(* IEC 61131-3 sources: plc-st-coding-agent/progress/evidence/f14_v3_parallel_20261112/jobs/codex_minimax-m27 (part 2) *)

(* ---- public-hard-05.raw_candidate_01.st ---- *)
FUNCTION_BLOCK MechanicalArmControl
VAR_INPUT
    ManualMode      : BOOL;
    SingleStepMode  : BOOL;
    SingleCycleMode : BOOL;
    ContinuousMode  : BOOL;
    EmergencyStop   : BOOL;
    Start           : BOOL;
    DownButton      : BOOL;
    UpButton        : BOOL;
    LeftButton      : BOOL;
    RightButton     : BOOL;
    GripButton      : BOOL;
    ReleaseButton   : BOOL;
    DownLimitSwitch     : BOOL;
    UpLimitSwitch       : BOOL;
    LeftLimitSwitch     : BOOL;
    RightLimitSwitch    : BOOL;
    GripLimitSwitch     : BOOL;
    ReleaseLimitSwitch  : BOOL;
END_VAR

VAR_OUTPUT
    MoveDown        : BOOL;
    MoveUp          : BOOL;
    MoveLeft        : BOOL;
    MoveRight       : BOOL;
    ActivateGrip    : BOOL;
    ActivateRelease : BOOL;
END_VAR

VAR
    stepNumber       : INT := 0;
    startRisingEdge  : BOOL;
    lastStart        : BOOL := FALSE;
    actionInProgress : BOOL := FALSE;
END_VAR

// Edge detection for Start button
startRisingEdge := Start AND NOT lastStart;
lastStart := Start;

// Emergency stop: highest priority, resets all outputs and state
IF NOT EmergencyStop THEN
    MoveDown        := FALSE;
    MoveUp          := FALSE;
    MoveLeft        := FALSE;
    MoveRight       := FALSE;
    ActivateGrip    := FALSE;
    ActivateRelease := FALSE;
    stepNumber      := 0;
    actionInProgress := FALSE;
ELSE
    // Manual mode control
    IF ManualMode THEN
        MoveDown        := DownButton AND NOT DownLimitSwitch;
        MoveUp          := UpButton AND NOT UpLimitSwitch;
        MoveLeft        := LeftButton AND NOT LeftLimitSwitch;
        MoveRight       := RightButton AND NOT RightLimitSwitch;
        ActivateGrip    := GripButton AND NOT GripLimitSwitch;
        ActivateRelease := ReleaseButton AND NOT ReleaseLimitSwitch;
        stepNumber      := 0;
        actionInProgress := FALSE;

    // Single step mode: Start button advances through steps
    ELSIF SingleStepMode THEN
        IF startRisingEdge AND NOT actionInProgress THEN
            stepNumber := stepNumber + 1;
        END_IF;

        CASE stepNumber OF
            1:
                MoveDown := TRUE;
                actionInProgress := TRUE;
                IF DownLimitSwitch THEN
                    MoveDown := FALSE;
                    actionInProgress := FALSE;
                END_IF;
            2:
                ActivateGrip := TRUE;
                actionInProgress := TRUE;
                IF GripLimitSwitch THEN
                    ActivateGrip := FALSE;
                    actionInProgress := FALSE;
                END_IF;
            3:
                MoveUp := TRUE;
                actionInProgress := TRUE;
                IF UpLimitSwitch THEN
                    MoveUp := FALSE;
                    actionInProgress := FALSE;
                END_IF;
            4:
                MoveRight := TRUE;
                actionInProgress := TRUE;
                IF RightLimitSwitch THEN
                    MoveRight := FALSE;
                    actionInProgress := FALSE;
                END_IF;
            5:
                MoveDown := TRUE;
                actionInProgress := TRUE;
                IF DownLimitSwitch THEN
                    MoveDown := FALSE;
                    actionInProgress := FALSE;
                END_IF;
            6:
                ActivateRelease := TRUE;
                actionInProgress := TRUE;
                IF ReleaseLimitSwitch THEN
                    ActivateRelease := FALSE;
                    actionInProgress := FALSE;
                END_IF;
            7:
                MoveUp := TRUE;
                actionInProgress := TRUE;
                IF UpLimitSwitch THEN
                    MoveUp := FALSE;
                    actionInProgress := FALSE;
                END_IF;
            8:
                MoveLeft := TRUE;
                actionInProgress := TRUE;
                IF LeftLimitSwitch THEN
                    MoveLeft := FALSE;
                    actionInProgress := FALSE;
                END_IF;
        END_CASE;

        IF stepNumber > 8 THEN
            stepNumber := 0;
        END_IF;

    // Single cycle mode: executes full cycle once then stops
    ELSIF SingleCycleMode THEN
        IF startRisingEdge THEN
            stepNumber := 1;
            actionInProgress := FALSE;
        END_IF;

        CASE stepNumber OF
            1:
                MoveDown := TRUE;
                actionInProgress := TRUE;
                IF DownLimitSwitch THEN
                    MoveDown := FALSE;
                    actionInProgress := FALSE;
                    stepNumber := 2;
                END_IF;
            2:
                ActivateGrip := TRUE;
                actionInProgress := TRUE;
                IF GripLimitSwitch THEN
                    ActivateGrip := FALSE;
                    actionInProgress := FALSE;
                    stepNumber := 3;
                END_IF;
            3:
                MoveUp := TRUE;
                actionInProgress := TRUE;
                IF UpLimitSwitch THEN
                    MoveUp := FALSE;
                    actionInProgress := FALSE;
                    stepNumber := 4;
                END_IF;
            4:
                MoveRight := TRUE;
                actionInProgress := TRUE;
                IF RightLimitSwitch THEN
                    MoveRight := FALSE;
                    actionInProgress := FALSE;
                    stepNumber := 5;
                END_IF;
            5:
                MoveDown := TRUE;
                actionInProgress := TRUE;
                IF DownLimitSwitch THEN
                    MoveDown := FALSE;
                    actionInProgress := FALSE;
                    stepNumber := 6;
                END_IF;
            6:
                ActivateRelease := TRUE;
                actionInProgress := TRUE;
                IF ReleaseLimitSwitch THEN
                    ActivateRelease := FALSE;
                    actionInProgress := FALSE;
                    stepNumber := 7;
                END_IF;
            7:
                MoveUp := TRUE;
                actionInProgress := TRUE;
                IF UpLimitSwitch THEN
                    MoveUp := FALSE;
                    actionInProgress := FALSE;
                    stepNumber := 8;
                END_IF;
            8:
                MoveLeft := TRUE;
                actionInProgress := TRUE;
                IF LeftLimitSwitch THEN
                    MoveLeft := FALSE;
                    actionInProgress := FALSE;
                    stepNumber := 0;
                END_IF;
        END_CASE;

    // Continuous mode: executes full cycle repeatedly
    ELSIF ContinuousMode THEN
        IF startRisingEdge THEN
            stepNumber := 1;
            actionInProgress := FALSE;
        END_IF;

        CASE stepNumber OF
            1:
                MoveDown := TRUE;
                actionInProgress := TRUE;
                IF DownLimitSwitch THEN
                    MoveDown := FALSE;
                    actionInProgress := FALSE;
                    stepNumber := 2;
                END_IF;
            2:
                ActivateGrip := TRUE;
                actionInProgress := TRUE;
                IF GripLimitSwitch THEN
                    ActivateGrip := FALSE;
                    actionInProgress := FALSE;
                    stepNumber := 3;
                END_IF;
            3:
                MoveUp := TRUE;
                actionInProgress := TRUE;
                IF UpLimitSwitch THEN
                    MoveUp := FALSE;
                    actionInProgress := FALSE;
                    stepNumber := 4;
                END_IF;
            4:
                MoveRight := TRUE;
                actionInProgress := TRUE;
                IF RightLimitSwitch THEN
                    MoveRight := FALSE;
                    actionInProgress := FALSE;
                    stepNumber := 5;
                END_IF;
            5:
                MoveDown := TRUE;
                actionInProgress := TRUE;
                IF DownLimitSwitch THEN
                    MoveDown := FALSE;
                    actionInProgress := FALSE;
                    stepNumber := 6;
                END_IF;
            6:
                ActivateRelease := TRUE;
                actionInProgress := TRUE;
                IF ReleaseLimitSwitch THEN
                    ActivateRelease := FALSE;
                    actionInProgress := FALSE;
                    stepNumber := 7;
                END_IF;
            7:
                MoveUp := TRUE;
                actionInProgress := TRUE;
                IF UpLimitSwitch THEN
                    MoveUp := FALSE;
                    actionInProgress := FALSE;
                    stepNumber := 8;
                END_IF;
            8:
                MoveLeft := TRUE;
                actionInProgress := TRUE;
                IF LeftLimitSwitch THEN
                    MoveLeft := FALSE;
                    actionInProgress := FALSE;
                    stepNumber := 1;
                END_IF;
        END_CASE;
    END_IF;
END_IF;
END_FUNCTION_BLOCK

(* ---- public-hard-05.raw_candidate_02.st ---- *)
FUNCTION_BLOCK MechanicalArmControl
VAR_INPUT
    ManualMode      : BOOL;
    SingleStepMode  : BOOL;
    SingleCycleMode : BOOL;
    ContinuousMode  : BOOL;
    EmergencyStop   : BOOL;
    Start           : BOOL;
    DownButton      : BOOL;
    UpButton        : BOOL;
    LeftButton      : BOOL;
    RightButton     : BOOL;
    GripButton      : BOOL;
    ReleaseButton   : BOOL;
    DownLimitSwitch     : BOOL;
    UpLimitSwitch       : BOOL;
    LeftLimitSwitch     : BOOL;
    RightLimitSwitch    : BOOL;
    GripLimitSwitch     : BOOL;
    ReleaseLimitSwitch  : BOOL;
END_VAR

VAR_OUTPUT
    MoveDown        : BOOL;
    MoveUp          : BOOL;
    MoveLeft        : BOOL;
    MoveRight       : BOOL;
    ActivateGrip    : BOOL;
    ActivateRelease : BOOL;
END_VAR

VAR
    stepNumber       : INT := 0;
    startRisingEdge  : BOOL;
    lastStart        : BOOL := FALSE;
    actionInProgress : BOOL := FALSE;
END_VAR

startRisingEdge := Start AND NOT lastStart;
lastStart := Start;

IF NOT EmergencyStop THEN
    MoveDown        := FALSE;
    MoveUp          := FALSE;
    MoveLeft        := FALSE;
    MoveRight       := FALSE;
    ActivateGrip    := FALSE;
    ActivateRelease := FALSE;
    stepNumber      := 0;
    actionInProgress := FALSE;
ELSE
    IF ManualMode THEN
        IF DownButton AND UpButton THEN
            MoveDown := FALSE;
            MoveUp := FALSE;
        ELSE
            MoveDown := DownButton AND NOT DownLimitSwitch;
            MoveUp := UpButton AND NOT UpLimitSwitch;
        END_IF;
        IF LeftButton AND RightButton THEN
            MoveLeft := FALSE;
            MoveRight := FALSE;
        ELSE
            MoveLeft := LeftButton AND NOT LeftLimitSwitch;
            MoveRight := RightButton AND NOT RightLimitSwitch;
        END_IF;
        ActivateGrip := GripButton AND NOT GripLimitSwitch;
        ActivateRelease := ReleaseButton AND NOT ReleaseLimitSwitch;
        stepNumber := 0;
        actionInProgress := FALSE;

    ELSIF SingleStepMode THEN
        IF startRisingEdge AND NOT actionInProgress THEN
            stepNumber := stepNumber + 1;
        END_IF;

        IF stepNumber = 0 THEN
            actionInProgress := FALSE;
        END_IF;

        CASE stepNumber OF
            1:
                MoveDown := TRUE;
                actionInProgress := TRUE;
                IF DownLimitSwitch THEN
                    MoveDown := FALSE;
                    actionInProgress := FALSE;
                END_IF;
            2:
                ActivateGrip := TRUE;
                actionInProgress := TRUE;
                IF GripLimitSwitch THEN
                    ActivateGrip := FALSE;
                    actionInProgress := FALSE;
                END_IF;
            3:
                MoveUp := TRUE;
                actionInProgress := TRUE;
                IF UpLimitSwitch THEN
                    MoveUp := FALSE;
                    actionInProgress := FALSE;
                END_IF;
            4:
                MoveRight := TRUE;
                actionInProgress := TRUE;
                IF RightLimitSwitch THEN
                    MoveRight := FALSE;
                    actionInProgress := FALSE;
                END_IF;
            5:
                MoveDown := TRUE;
                actionInProgress := TRUE;
                IF DownLimitSwitch THEN
                    MoveDown := FALSE;
                    actionInProgress := FALSE;
                END_IF;
            6:
                ActivateRelease := TRUE;
                actionInProgress := TRUE;
                IF ReleaseLimitSwitch THEN
                    ActivateRelease := FALSE;
                    actionInProgress := FALSE;
                END_IF;
            7:
                MoveUp := TRUE;
                actionInProgress := TRUE;
                IF UpLimitSwitch THEN
                    MoveUp := FALSE;
                    actionInProgress := FALSE;
                END_IF;
            8:
                MoveLeft := TRUE;
                actionInProgress := TRUE;
                IF LeftLimitSwitch THEN
                    MoveLeft := FALSE;
                    actionInProgress := FALSE;
                END_IF;
        END_CASE;

        IF stepNumber > 8 THEN
            stepNumber := 0;
        END_IF;

    ELSIF SingleCycleMode THEN
        IF startRisingEdge THEN
            stepNumber := 1;
            actionInProgress := FALSE;
        END_IF;

        IF stepNumber = 0 THEN
            actionInProgress := FALSE;
        END_IF;

        CASE stepNumber OF
            1:
                MoveDown := TRUE;
                actionInProgress := TRUE;
                IF DownLimitSwitch THEN
                    MoveDown := FALSE;
                    actionInProgress := FALSE;
                    stepNumber := 2;
                END_IF;
            2:
                ActivateGrip := TRUE;
                actionInProgress := TRUE;
                IF GripLimitSwitch THEN
                    ActivateGrip := FALSE;
                    actionInProgress := FALSE;
                    stepNumber := 3;
                END_IF;
            3:
                MoveUp := TRUE;
                actionInProgress := TRUE;
                IF UpLimitSwitch THEN
                    MoveUp := FALSE;
                    actionInProgress := FALSE;
                    stepNumber := 4;
                END_IF;
            4:
                MoveRight := TRUE;
                actionInProgress := TRUE;
                IF RightLimitSwitch THEN
                    MoveRight := FALSE;
                    actionInProgress := FALSE;
                    stepNumber := 5;
                END_IF;
            5:
                MoveDown := TRUE;
                actionInProgress := TRUE;
                IF DownLimitSwitch THEN
                    MoveDown := FALSE;
                    actionInProgress := FALSE;
                    stepNumber := 6;
                END_IF;
            6:
                ActivateRelease := TRUE;
                actionInProgress := TRUE;
                IF ReleaseLimitSwitch THEN
                    ActivateRelease := FALSE;
                    actionInProgress := FALSE;
                    stepNumber := 7;
                END_IF;
            7:
                MoveUp := TRUE;
                actionInProgress := TRUE;
                IF UpLimitSwitch THEN
                    MoveUp := FALSE;
                    actionInProgress := FALSE;
                    stepNumber := 8;
                END_IF;
            8:
                MoveLeft := TRUE;
                actionInProgress := TRUE;
                IF LeftLimitSwitch THEN
                    MoveLeft := FALSE;
                    actionInProgress := FALSE;
                    stepNumber := 0;
                END_IF;
        END_CASE;

    ELSIF ContinuousMode THEN
        IF startRisingEdge THEN
            stepNumber := 1;
            actionInProgress := FALSE;
        END_IF;

        IF stepNumber = 0 THEN
            actionInProgress := FALSE;
        END_IF;

        CASE stepNumber OF
            1:
                MoveDown := TRUE;
                actionInProgress := TRUE;
                IF DownLimitSwitch THEN
                    MoveDown := FALSE;
                    actionInProgress := FALSE;
                    stepNumber := 2;
                END_IF;
            2:
                ActivateGrip := TRUE;
                actionInProgress := TRUE;
                IF GripLimitSwitch THEN
                    ActivateGrip := FALSE;
                    actionInProgress := FALSE;
                    stepNumber := 3;
                END_IF;
            3:
                MoveUp := TRUE;
                actionInProgress := TRUE;
                IF UpLimitSwitch THEN
                    MoveUp := FALSE;
                    actionInProgress := FALSE;
                    stepNumber := 4;
                END_IF;
            4:
                MoveRight := TRUE;
                actionInProgress := TRUE;
                IF RightLimitSwitch THEN
                    MoveRight := FALSE;
                    actionInProgress := FALSE;
                    stepNumber := 5;
                END_IF;
            5:
                MoveDown := TRUE;
                actionInProgress := TRUE;
                IF DownLimitSwitch THEN
                    MoveDown := FALSE;
                    actionInProgress := FALSE;
                    stepNumber := 6;
                END_IF;
            6:
                ActivateRelease := TRUE;
                actionInProgress := TRUE;
                IF ReleaseLimitSwitch THEN
                    ActivateRelease := FALSE;
                    actionInProgress := FALSE;
                    stepNumber := 7;
                END_IF;
            7:
                MoveUp := TRUE;
                actionInProgress := TRUE;
                IF UpLimitSwitch THEN
                    MoveUp := FALSE;
                    actionInProgress := FALSE;
                    stepNumber := 8;
                END_IF;
            8:
                MoveLeft := TRUE;
                actionInProgress := TRUE;
                IF LeftLimitSwitch THEN
                    MoveLeft := FALSE;
                    actionInProgress := FALSE;
                    stepNumber := 1;
                END_IF;
        END_CASE;
    END_IF;
END_IF;
END_FUNCTION_BLOCK

(* ---- public-hard-06.candidate_01.st ---- *)
TYPE ProductState : (
    Idle := 0,
    AtFeed := 1,
    AtWash := 2,
    AtWeight := 3,
    AtFiring := 4,
    AtOutput := 5,
    Rejected := 6
);
END_TYPE;

FUNCTION_BLOCK ProductionControl
VAR_INPUT
    Mode : BOOL;
    ForwardButton : BOOL;
    ReverseButton : BOOL;
    SensorFeed : BOOL;
    SensorWash : BOOL;
    SensorWeight : BOOL;
    SensorFiring : BOOL;
    SensorOutput : BOOL;
    washComplete : BOOL;
    weightComplete : BOOL;
    weight : REAL;
    firingComplete : BOOL;
END_VAR

VAR_OUTPUT
    MotorForward : BOOL := FALSE;
    MotorReverse : BOOL := FALSE;
    kick : BOOL := FALSE;
    CompletionLight : BOOL := FALSE;
    firingTemp : REAL := 0.0;
END_VAR

VAR
    currentState : ProductState := Idle;
    prevSensorFeed : BOOL := FALSE;
    prevSensorWash : BOOL := FALSE;
    prevSensorWeight : BOOL := FALSE;
    prevSensorFiring : BOOL := FALSE;
    prevSensorOutput : BOOL := FALSE;
END_VAR

IF currentState = Idle THEN
    MotorForward := FALSE;
    MotorReverse := FALSE;
    kick := FALSE;
    CompletionLight := FALSE;
    firingTemp := 0.0;
END_IF;

IF Mode = FALSE THEN
    MotorForward := ForwardButton;
    MotorReverse := ReverseButton AND NOT ForwardButton;
    MotorReverse := MotorReverse;
ELSE
    MotorReverse := FALSE;

    IF currentState = Idle THEN
        IF SensorFeed AND NOT prevSensorFeed THEN
            currentState := AtFeed;
            MotorForward := TRUE;
        END_IF;

    ELSIF currentState = AtFeed THEN
        MotorForward := TRUE;
        IF SensorWash AND NOT prevSensorWash THEN
            currentState := AtWash;
            MotorForward := FALSE;
        END_IF;

    ELSIF currentState = AtWash THEN
        MotorForward := FALSE;
        IF washComplete THEN
            currentState := AtWeight;
            MotorForward := TRUE;
        END_IF;

    ELSIF currentState = AtWeight THEN
        MotorForward := FALSE;
        IF weightComplete THEN
            IF weight < 100.0 OR weight > 200.0 THEN
                kick := TRUE;
                currentState := Rejected;
                MotorForward := TRUE;
            ELSE
                firingTemp := 500.0 + (weight - 100.0) * 0.5;
                currentState := AtFiring;
                MotorForward := TRUE;
            END_IF;
        END_IF;

    ELSIF currentState = AtFiring THEN
        MotorForward := FALSE;
        IF firingComplete THEN
            currentState := AtOutput;
            MotorForward := FALSE;
            CompletionLight := TRUE;
        END_IF;

    ELSIF currentState = AtOutput THEN
        MotorForward := FALSE;
        CompletionLight := SensorOutput;
        IF NOT SensorOutput AND prevSensorOutput THEN
            currentState := Idle;
            CompletionLight := FALSE;
        END_IF;

    ELSIF currentState = Rejected THEN
        MotorForward := TRUE;
        kick := SensorWeight;
        IF NOT SensorWeight AND prevSensorWeight THEN
            currentState := Idle;
            kick := FALSE;
        END_IF;

    END_IF;
END_IF;

prevSensorFeed := SensorFeed;
prevSensorWash := SensorWash;
prevSensorWeight := SensorWeight;
prevSensorFiring := SensorFiring;
prevSensorOutput := SensorOutput;

END_FUNCTION_BLOCK

(* ---- public-hard-06.candidate_02.st ---- *)
TYPE ProductState : (
    Idle := 0,
    AtFeed := 1,
    AtWash := 2,
    AtWeight := 3,
    AtFiring := 4,
    AtOutput := 5,
    Rejected := 6
);
END_TYPE;

TYPE ModeType : (Manual := 0, Auto := 1, Sequence := 2);
END_TYPE;

FUNCTION_BLOCK ProductionControl
VAR_INPUT
    Mode : BOOL;
    ForwardButton : BOOL;
    ReverseButton : BOOL;
    SensorFeed : BOOL;
    SensorWash : BOOL;
    SensorWeight : BOOL;
    SensorFiring : BOOL;
    SensorOutput : BOOL;
    washComplete : BOOL;
    weightComplete : BOOL;
    weight : REAL;
    firingComplete : BOOL;
END_VAR

VAR_OUTPUT
    MotorForward : BOOL := FALSE;
    MotorReverse : BOOL := FALSE;
    kick : BOOL := FALSE;
    CompletionLight : BOOL := FALSE;
    firingTemp : REAL := 0.0;
END_VAR

VAR
    currentState : ProductState := Idle;
    prevSensorFeed : BOOL := FALSE;
    prevSensorWash : BOOL := FALSE;
    prevSensorWeight : BOOL := FALSE;
    prevSensorFiring : BOOL := FALSE;
    prevSensorOutput : BOOL := FALSE;
    prevWashComplete : BOOL := FALSE;
    prevWeightComplete : BOOL := FALSE;
    prevFiringComplete : BOOL := FALSE;
END_VAR

IF currentState = Idle THEN
    MotorForward := FALSE;
    MotorReverse := FALSE;
    kick := FALSE;
    CompletionLight := FALSE;
    firingTemp := 0.0;
END_IF;

IF Mode = FALSE THEN
    MotorForward := ForwardButton;
    MotorReverse := ReverseButton AND NOT ForwardButton;
ELSE
    MotorReverse := FALSE;

    IF currentState = Idle THEN
        IF SensorFeed AND NOT prevSensorFeed THEN
            currentState := AtFeed;
            MotorForward := TRUE;
        END_IF;

    ELSIF currentState = AtFeed THEN
        MotorForward := TRUE;
        IF SensorWash AND NOT prevSensorWash THEN
            currentState := AtWash;
            MotorForward := FALSE;
        END_IF;

    ELSIF currentState = AtWash THEN
        MotorForward := FALSE;
        IF washComplete AND NOT prevWashComplete THEN
            currentState := AtWeight;
            MotorForward := TRUE;
        END_IF;

    ELSIF currentState = AtWeight THEN
        MotorForward := FALSE;
        IF weightComplete AND NOT prevWeightComplete THEN
            IF weight < 100.0 OR weight > 200.0 THEN
                kick := TRUE;
                currentState := Rejected;
            ELSE
                firingTemp := 500.0 + (weight - 100.0) * 0.5;
                currentState := AtFiring;
            END_IF;
        END_IF;

    ELSIF currentState = AtFiring THEN
        MotorForward := FALSE;
        IF firingComplete AND NOT prevFiringComplete THEN
            currentState := AtOutput;
            CompletionLight := TRUE;
        END_IF;

    ELSIF currentState = AtOutput THEN
        MotorForward := FALSE;
        CompletionLight := SensorOutput;
        IF NOT SensorOutput AND prevSensorOutput THEN
            currentState := Idle;
            CompletionLight := FALSE;
        END_IF;

    ELSIF currentState = Rejected THEN
        MotorForward := FALSE;
        kick := SensorWeight;
        IF NOT SensorWeight AND prevSensorWeight THEN
            currentState := Idle;
            kick := FALSE;
        END_IF;

    END_IF;
END_IF;

prevSensorFeed := SensorFeed;
prevSensorWash := SensorWash;
prevSensorWeight := SensorWeight;
prevSensorFiring := SensorFiring;
prevSensorOutput := SensorOutput;
prevWashComplete := washComplete;
prevWeightComplete := weightComplete;
prevFiringComplete := firingComplete;

END_FUNCTION_BLOCK

(* ---- public-hard-06.raw_candidate_01.st ---- *)
TYPE ProductState : (
    Idle := 0,
    AtFeed := 1,
    AtWash := 2,
    AtWeight := 3,
    AtFiring := 4,
    AtOutput := 5,
    Rejected := 6
);
END_TYPE

FUNCTION_BLOCK ProductionControl
VAR_INPUT
    Mode : BOOL;
    ForwardButton : BOOL;
    ReverseButton : BOOL;
    SensorFeed : BOOL;
    SensorWash : BOOL;
    SensorWeight : BOOL;
    SensorFiring : BOOL;
    SensorOutput : BOOL;
    washComplete : BOOL;
    weightComplete : BOOL;
    weight : REAL;
    firingComplete : BOOL;
END_VAR

VAR_OUTPUT
    MotorForward : BOOL := FALSE;
    MotorReverse : BOOL := FALSE;
    kick : BOOL := FALSE;
    CompletionLight : BOOL := FALSE;
    firingTemp : REAL := 0.0;
END_VAR

VAR
    currentState : ProductState := Idle;
    prevSensorFeed : BOOL := FALSE;
    prevSensorWash : BOOL := FALSE;
    prevSensorWeight : BOOL := FALSE;
    prevSensorFiring : BOOL := FALSE;
    prevSensorOutput : BOOL := FALSE;
END_VAR

IF currentState = Idle THEN
    MotorForward := FALSE;
    MotorReverse := FALSE;
    kick := FALSE;
    CompletionLight := FALSE;
    firingTemp := 0.0;
END_IF

IF Mode = FALSE THEN
    MotorForward := ForwardButton;
    MotorReverse := ReverseButton AND NOT ForwardButton;
    MotorReverse := MotorReverse;
ELSE
    MotorReverse := FALSE;

    IF currentState = Idle THEN
        IF SensorFeed AND NOT prevSensorFeed THEN
            currentState := AtFeed;
            MotorForward := TRUE;
        END_IF

    ELSIF currentState = AtFeed THEN
        MotorForward := TRUE;
        IF SensorWash AND NOT prevSensorWash THEN
            currentState := AtWash;
            MotorForward := FALSE;
        END_IF

    ELSIF currentState = AtWash THEN
        MotorForward := FALSE;
        IF washComplete THEN
            currentState := AtWeight;
            MotorForward := TRUE;
        END_IF

    ELSIF currentState = AtWeight THEN
        MotorForward := FALSE;
        IF weightComplete THEN
            IF weight < 100.0 OR weight > 200.0 THEN
                kick := TRUE;
                currentState := Rejected;
                MotorForward := TRUE;
            ELSE
                firingTemp := 500.0 + (weight - 100.0) * 0.5;
                currentState := AtFiring;
                MotorForward := TRUE;
            END_IF;
        END_IF

    ELSIF currentState = AtFiring THEN
        MotorForward := FALSE;
        IF firingComplete THEN
            currentState := AtOutput;
            MotorForward := FALSE;
            CompletionLight := TRUE;
        END_IF

    ELSIF currentState = AtOutput THEN
        MotorForward := FALSE;
        CompletionLight := SensorOutput;
        IF NOT SensorOutput AND prevSensorOutput THEN
            currentState := Idle;
            CompletionLight := FALSE;
        END_IF

    ELSIF currentState = Rejected THEN
        MotorForward := TRUE;
        kick := SensorWeight;
        IF NOT SensorWeight AND prevSensorWeight THEN
            currentState := Idle;
            kick := FALSE;
        END_IF

    END_IF
END_IF

prevSensorFeed := SensorFeed;
prevSensorWash := SensorWash;
prevSensorWeight := SensorWeight;
prevSensorFiring := SensorFiring;
prevSensorOutput := SensorOutput;

END_FUNCTION_BLOCK

(* ---- public-hard-06.raw_candidate_02.st ---- *)
TYPE ProductState : (
    Idle := 0,
    AtFeed := 1,
    AtWash := 2,
    AtWeight := 3,
    AtFiring := 4,
    AtOutput := 5,
    Rejected := 6
);
END_TYPE

TYPE ModeType : (Manual := 0, Auto := 1, Sequence := 2);
END_TYPE

FUNCTION_BLOCK ProductionControl
VAR_INPUT
    Mode : BOOL;
    ForwardButton : BOOL;
    ReverseButton : BOOL;
    SensorFeed : BOOL;
    SensorWash : BOOL;
    SensorWeight : BOOL;
    SensorFiring : BOOL;
    SensorOutput : BOOL;
    washComplete : BOOL;
    weightComplete : BOOL;
    weight : REAL;
    firingComplete : BOOL;
END_VAR

VAR_OUTPUT
    MotorForward : BOOL := FALSE;
    MotorReverse : BOOL := FALSE;
    kick : BOOL := FALSE;
    CompletionLight : BOOL := FALSE;
    firingTemp : REAL := 0.0;
END_VAR

VAR
    currentState : ProductState := Idle;
    prevSensorFeed : BOOL := FALSE;
    prevSensorWash : BOOL := FALSE;
    prevSensorWeight : BOOL := FALSE;
    prevSensorFiring : BOOL := FALSE;
    prevSensorOutput : BOOL := FALSE;
    prevWashComplete : BOOL := FALSE;
    prevWeightComplete : BOOL := FALSE;
    prevFiringComplete : BOOL := FALSE;
END_VAR

IF currentState = Idle THEN
    MotorForward := FALSE;
    MotorReverse := FALSE;
    kick := FALSE;
    CompletionLight := FALSE;
    firingTemp := 0.0;
END_IF;

IF Mode = FALSE THEN
    MotorForward := ForwardButton;
    MotorReverse := ReverseButton AND NOT ForwardButton;
ELSE
    MotorReverse := FALSE;

    IF currentState = Idle THEN
        IF SensorFeed AND NOT prevSensorFeed THEN
            currentState := AtFeed;
            MotorForward := TRUE;
        END_IF;

    ELSIF currentState = AtFeed THEN
        MotorForward := TRUE;
        IF SensorWash AND NOT prevSensorWash THEN
            currentState := AtWash;
            MotorForward := FALSE;
        END_IF;

    ELSIF currentState = AtWash THEN
        MotorForward := FALSE;
        IF washComplete AND NOT prevWashComplete THEN
            currentState := AtWeight;
            MotorForward := TRUE;
        END_IF;

    ELSIF currentState = AtWeight THEN
        MotorForward := FALSE;
        IF weightComplete AND NOT prevWeightComplete THEN
            IF weight < 100.0 OR weight > 200.0 THEN
                kick := TRUE;
                currentState := Rejected;
            ELSE
                firingTemp := 500.0 + (weight - 100.0) * 0.5;
                currentState := AtFiring;
            END_IF;
        END_IF;

    ELSIF currentState = AtFiring THEN
        MotorForward := FALSE;
        IF firingComplete AND NOT prevFiringComplete THEN
            currentState := AtOutput;
            CompletionLight := TRUE;
        END_IF;

    ELSIF currentState = AtOutput THEN
        MotorForward := FALSE;
        CompletionLight := SensorOutput;
        IF NOT SensorOutput AND prevSensorOutput THEN
            currentState := Idle;
            CompletionLight := FALSE;
        END_IF;

    ELSIF currentState = Rejected THEN
        MotorForward := FALSE;
        kick := SensorWeight;
        IF NOT SensorWeight AND prevSensorWeight THEN
            currentState := Idle;
            kick := FALSE;
        END_IF;

    END_IF;
END_IF;

prevSensorFeed := SensorFeed;
prevSensorWash := SensorWash;
prevSensorWeight := SensorWeight;
prevSensorFiring := SensorFiring;
prevSensorOutput := SensorOutput;
prevWashComplete := washComplete;
prevWeightComplete := weightComplete;
prevFiringComplete := firingComplete;

END_FUNCTION_BLOCK

(* ---- public-medium-01.candidate_01.st ---- *)
FUNCTION_BLOCK FB_PumpControl
VAR
    i : INT;
    sortedIndices : ARRAY[1..5] OF INT;
    temp : INT;
    j : INT;
END_VAR

    // Stop button has highest priority
    IF stop THEN
        FOR i := 1 TO 5 DO
            pumpGroup[i].RunComd := FALSE;
        END_FOR;
        RETURN;
    END_IF;

    // Start button applies mode-specific logic
    IF start THEN
        IF NOT mode THEN
            // Manual mode - run pumps where selection is TRUE
            FOR i := 1 TO 5 DO
                pumpGroup[i].RunComd := pumpGroup[i].selection;
            END_FOR;
        ELSE
            // Automatic mode - select 3 pumps with highest priority
            FOR i := 1 TO 5 DO
                sortedIndices[i] := i;
            END_FOR;

            // Bubble sort by priority (descending)
            FOR i := 1 TO 4 DO
                FOR j := i + 1 TO 5 DO
                    IF pumpGroup[sortedIndices[j]].priority > pumpGroup[sortedIndices[i]].priority THEN
                        temp := sortedIndices[i];
                        sortedIndices[i] := sortedIndices[j];
                        sortedIndices[j] := temp;
                    END_IF;
                END_FOR;
            END_FOR;

            // Deactivate all pumps first
            FOR i := 1 TO 5 DO
                pumpGroup[i].RunComd := FALSE;
            END_FOR;

            // Activate top 3 pumps by priority
            FOR i := 1 TO 3 DO
                pumpGroup[sortedIndices[i]].RunComd := TRUE;
            END_FOR;
        END_IF;
    END_IF;
END_FUNCTION_BLOCK

(* ---- public-medium-01.candidate_02.st ---- *)
TYPE ST_Pump :
STRUCT
    priority : INT;
    selection : BOOL;
    RunComd : BOOL;
END_STRUCT;
END_TYPE;

FUNCTION_BLOCK FB_PumpControl
VAR_INPUT
    mode : BOOL;
    start : BOOL;
    stop : BOOL;
END_VAR

VAR_IN_OUT
    pumpGroup : ARRAY[1..5] OF ST_Pump;
END_VAR

VAR
    i : INT;
    sortedIndices : ARRAY[1..5] OF INT;
    temp : INT;
    j : INT;
END_VAR

    IF stop THEN
        FOR i := 1 TO 5 DO
            pumpGroup[i].RunComd := FALSE;
        END_FOR;
        RETURN;
    END_IF;

    IF start THEN
        IF NOT mode THEN
            FOR i := 1 TO 5 DO
                pumpGroup[i].RunComd := pumpGroup[i].selection;
            END_FOR;
        ELSE
            FOR i := 1 TO 5 DO
                sortedIndices[i] := i;
            END_FOR;

            FOR i := 1 TO 4 DO
                FOR j := i + 1 TO 5 DO
                    IF pumpGroup[sortedIndices[j]].priority > pumpGroup[sortedIndices[i]].priority THEN
                        temp := sortedIndices[i];
                        sortedIndices[i] := sortedIndices[j];
                        sortedIndices[j] := temp;
                    END_IF;
                END_FOR;
            END_FOR;

            FOR i := 1 TO 5 DO
                pumpGroup[i].RunComd := FALSE;
            END_FOR;

            FOR i := 1 TO 3 DO
                pumpGroup[sortedIndices[i]].RunComd := TRUE;
            END_FOR;
        END_IF;
    END_IF;
END_FUNCTION_BLOCK

(* ---- public-medium-01.raw_candidate_01.st ---- *)
FUNCTION_BLOCK FB_PumpControl
VAR
    i : INT;
    sortedIndices : ARRAY[1..5] OF INT;
    temp : INT;
    j : INT;
END_VAR

    // Stop button has highest priority
    IF stop THEN
        FOR i := 1 TO 5 DO
            pumpGroup[i].RunComd := FALSE;
        END_FOR;
        RETURN;
    END_IF;

    // Start button applies mode-specific logic
    IF start THEN
        IF NOT mode THEN
            // Manual mode - run pumps where selection is TRUE
            FOR i := 1 TO 5 DO
                pumpGroup[i].RunComd := pumpGroup[i].selection;
            END_FOR;
        ELSE
            // Automatic mode - select 3 pumps with highest priority
            FOR i := 1 TO 5 DO
                sortedIndices[i] := i;
            END_FOR;

            // Bubble sort by priority (descending)
            FOR i := 1 TO 4 DO
                FOR j := i + 1 TO 5 DO
                    IF pumpGroup[sortedIndices[j]].priority > pumpGroup[sortedIndices[i]].priority THEN
                        temp := sortedIndices[i];
                        sortedIndices[i] := sortedIndices[j];
                        sortedIndices[j] := temp;
                    END_IF;
                END_FOR;
            END_FOR;

            // Deactivate all pumps first
            FOR i := 1 TO 5 DO
                pumpGroup[i].RunComd := FALSE;
            END_FOR;

            // Activate top 3 pumps by priority
            FOR i := 1 TO 3 DO
                pumpGroup[sortedIndices[i]].RunComd := TRUE;
            END_FOR;
        END_IF;
    END_IF;
END_FUNCTION_BLOCK

(* ---- public-medium-01.raw_candidate_02.st ---- *)
TYPE ST_Pump :
STRUCT
    priority : INT;
    selection : BOOL;
    RunComd : BOOL;
END_STRUCT
END_TYPE

FUNCTION_BLOCK FB_PumpControl
VAR_INPUT
    mode : BOOL;
    start : BOOL;
    stop : BOOL;
END_VAR

VAR_IN_OUT
    pumpGroup : ARRAY[1..5] OF ST_Pump;
END_VAR

VAR
    i : INT;
    sortedIndices : ARRAY[1..5] OF INT;
    temp : INT;
    j : INT;
END_VAR

    IF stop THEN
        FOR i := 1 TO 5 DO
            pumpGroup[i].RunComd := FALSE;
        END_FOR;
        RETURN;
    END_IF;

    IF start THEN
        IF NOT mode THEN
            FOR i := 1 TO 5 DO
                pumpGroup[i].RunComd := pumpGroup[i].selection;
            END_FOR;
        ELSE
            FOR i := 1 TO 5 DO
                sortedIndices[i] := i;
            END_FOR;

            FOR i := 1 TO 4 DO
                FOR j := i + 1 TO 5 DO
                    IF pumpGroup[sortedIndices[j]].priority > pumpGroup[sortedIndices[i]].priority THEN
                        temp := sortedIndices[i];
                        sortedIndices[i] := sortedIndices[j];
                        sortedIndices[j] := temp;
                    END_IF;
                END_FOR;
            END_FOR;

            FOR i := 1 TO 5 DO
                pumpGroup[i].RunComd := FALSE;
            END_FOR;

            FOR i := 1 TO 3 DO
                pumpGroup[sortedIndices[i]].RunComd := TRUE;
            END_FOR;
        END_IF;
    END_IF;
END_FUNCTION_BLOCK

(* ---- public-medium-02.candidate_01.st ---- *)
TYPE ST_AnalogChannel
STRUCT
    enable        : BOOL;
    hiLIM         : REAL;
    loLIM         : REAL;
    bipolar       : BOOL;
    measuringMode : INT;
    retVal        : WORD;
    outputValue   : REAL;
END_STRUCT;
END_TYPE;

FUNCTION_BLOCK FB_AnalogBatchProcessing
VAR_INPUT
    count : DINT;
END_VAR
VAR_IN_OUT
    analogValues : ARRAY[*] OF INT;
    channels     : ARRAY[*] OF ST_AnalogChannel;
END_VAR
VAR
    i         : DINT;
    lowerIdx  : DINT;
    upperIdx  : DINT;
    rawValue  : INT;
END_VAR

lowerIdx := LOWER_BOUND(analogValues, 1);
upperIdx := lowerIdx + count - 1;

FOR i := lowerIdx TO upperIdx DO
    rawValue := analogValues[i];

    IF channels[i].enable THEN
        CASE channels[i].measuringMode OF
            0: // Non-temperature linear scaling
                IF channels[i].hiLIM > channels[i].loLIM THEN
                    IF channels[i].bipolar THEN
                        channels[i].outputValue := channels[i].loLIM +
                            ((TO_REAL(rawValue) + 27648.0) / 55296.0) *
                            (channels[i].hiLIM - channels[i].loLIM);
                    ELSE
                        channels[i].outputValue := channels[i].loLIM +
                            (TO_REAL(rawValue) / 27648.0) *
                            (channels[i].hiLIM - channels[i].loLIM);
                    END_IF;
                    channels[i].retVal := 16#0000;
                ELSE
                    channels[i].retVal := 16#8002;
                END_IF;

            1: // Standard temperature
                channels[i].outputValue := TO_REAL(rawValue) / 10.0;
                channels[i].retVal := 16#0000;

            2: // Climatic temperature
                channels[i].outputValue := TO_REAL(rawValue) / 100.0;
                channels[i].retVal := 16#0000;

            ELSE
                channels[i].retVal := 16#8001;
        END_CASE;
    END_IF;
END_FOR;

END_FUNCTION_BLOCK

(* ---- public-medium-02.candidate_02.st ---- *)
TYPE ST_AnalogChannel :
STRUCT
    enable        : BOOL;
    hiLIM         : REAL;
    loLIM         : REAL;
    bipolar       : BOOL;
    measuringMode : INT;
    retVal        : WORD;
    outputValue   : REAL;
END_STRUCT;
END_TYPE;

FUNCTION_BLOCK FB_AnalogBatchProcessing
VAR_INPUT
    count : DINT;
END_VAR
VAR_IN_OUT
    analogValues : ARRAY[*] OF INT;
    channels     : ARRAY[*] OF ST_AnalogChannel;
END_VAR
VAR
    i         : DINT;
    lowerIdx  : DINT;
    upperIdx  : DINT;
    rawValue  : INT;
END_VAR

lowerIdx := LOWER_BOUND(analogValues, 1);
upperIdx := lowerIdx + count - 1;

FOR i := lowerIdx TO upperIdx DO
    rawValue := analogValues[i];

    IF channels[i].enable THEN
        CASE channels[i].measuringMode OF
            0: // Non-temperature linear scaling
                IF channels[i].hiLIM > channels[i].loLIM THEN
                    IF channels[i].bipolar THEN
                        channels[i].outputValue := channels[i].loLIM +
                            ((INT_TO_REAL(rawValue) + 27648.0) / 55296.0) *
                            (channels[i].hiLIM - channels[i].loLIM);
                    ELSE
                        channels[i].outputValue := channels[i].loLIM +
                            (INT_TO_REAL(rawValue) / 27648.0) *
                            (channels[i].hiLIM - channels[i].loLIM);
                    END_IF;
                    channels[i].retVal := 16#0000;
                ELSE
                    channels[i].retVal := 16#8002;
                END_IF;

            1: // Standard temperature
                channels[i].outputValue := INT_TO_REAL(rawValue) / 10.0;
                channels[i].retVal := 16#0000;

            2: // Climatic temperature
                channels[i].outputValue := INT_TO_REAL(rawValue) / 100.0;
                channels[i].retVal := 16#0000;

            ELSE
                channels[i].retVal := 16#8001;
        END_CASE;
    END_IF;
END_FOR;

END_FUNCTION_BLOCK

(* ---- public-medium-02.raw_candidate_01.st ---- *)
TYPE ST_AnalogChannel
STRUCT
    enable        : BOOL;
    hiLIM         : REAL;
    loLIM         : REAL;
    bipolar       : BOOL;
    measuringMode : INT;
    retVal        : WORD;
    outputValue   : REAL;
END_STRUCT
END_TYPE

FUNCTION_BLOCK FB_AnalogBatchProcessing
VAR_INPUT
    count : DINT;
END_VAR
VAR_IN_OUT
    analogValues : ARRAY[*] OF INT;
    channels     : ARRAY[*] OF ST_AnalogChannel;
END_VAR
VAR
    i         : DINT;
    lowerIdx  : DINT;
    upperIdx  : DINT;
    rawValue  : INT;
END_VAR

lowerIdx := LOWER_BOUND(analogValues, 1);
upperIdx := lowerIdx + count - 1;

FOR i := lowerIdx TO upperIdx DO
    rawValue := analogValues[i];

    IF channels[i].enable THEN
        CASE channels[i].measuringMode OF
            0: // Non-temperature linear scaling
                IF channels[i].hiLIM > channels[i].loLIM THEN
                    IF channels[i].bipolar THEN
                        channels[i].outputValue := channels[i].loLIM +
                            ((TO_REAL(rawValue) + 27648.0) / 55296.0) *
                            (channels[i].hiLIM - channels[i].loLIM);
                    ELSE
                        channels[i].outputValue := channels[i].loLIM +
                            (TO_REAL(rawValue) / 27648.0) *
                            (channels[i].hiLIM - channels[i].loLIM);
                    END_IF;
                    channels[i].retVal := 16#0000;
                ELSE
                    channels[i].retVal := 16#8002;
                END_IF;

            1: // Standard temperature
                channels[i].outputValue := TO_REAL(rawValue) / 10.0;
                channels[i].retVal := 16#0000;

            2: // Climatic temperature
                channels[i].outputValue := TO_REAL(rawValue) / 100.0;
                channels[i].retVal := 16#0000;

            ELSE
                channels[i].retVal := 16#8001;
        END_CASE;
    END_IF;
END_FOR;

END_FUNCTION_BLOCK

(* ---- public-medium-02.raw_candidate_02.st ---- *)
TYPE ST_AnalogChannel :
STRUCT
    enable        : BOOL;
    hiLIM         : REAL;
    loLIM         : REAL;
    bipolar       : BOOL;
    measuringMode : INT;
    retVal        : WORD;
    outputValue   : REAL;
END_STRUCT
END_TYPE

FUNCTION_BLOCK FB_AnalogBatchProcessing
VAR_INPUT
    count : DINT;
END_VAR
VAR_IN_OUT
    analogValues : ARRAY[*] OF INT;
    channels     : ARRAY[*] OF ST_AnalogChannel;
END_VAR
VAR
    i         : DINT;
    lowerIdx  : DINT;
    upperIdx  : DINT;
    rawValue  : INT;
END_VAR

lowerIdx := LOWER_BOUND(analogValues, 1);
upperIdx := lowerIdx + count - 1;

FOR i := lowerIdx TO upperIdx DO
    rawValue := analogValues[i];

    IF channels[i].enable THEN
        CASE channels[i].measuringMode OF
            0: // Non-temperature linear scaling
                IF channels[i].hiLIM > channels[i].loLIM THEN
                    IF channels[i].bipolar THEN
                        channels[i].outputValue := channels[i].loLIM +
                            ((INT_TO_REAL(rawValue) + 27648.0) / 55296.0) *
                            (channels[i].hiLIM - channels[i].loLIM);
                    ELSE
                        channels[i].outputValue := channels[i].loLIM +
                            (INT_TO_REAL(rawValue) / 27648.0) *
                            (channels[i].hiLIM - channels[i].loLIM);
                    END_IF;
                    channels[i].retVal := 16#0000;
                ELSE
                    channels[i].retVal := 16#8002;
                END_IF;

            1: // Standard temperature
                channels[i].outputValue := INT_TO_REAL(rawValue) / 10.0;
                channels[i].retVal := 16#0000;

            2: // Climatic temperature
                channels[i].outputValue := INT_TO_REAL(rawValue) / 100.0;
                channels[i].retVal := 16#0000;

            ELSE
                channels[i].retVal := 16#8001;
        END_CASE;
    END_IF;
END_FOR;

END_FUNCTION_BLOCK

(* ---- public-medium-03.candidate_01.st ---- *)
FUNCTION_BLOCK FB_MovingAverage
VAR_INPUT
    cyclicExecution : BOOL;
    trigger : BOOL;
    value : LREAL;
    windowSize : INT;
    reset : BOOL;
END_VAR

VAR_OUTPUT
    average : LREAL := 0.0;
    windowSizeReached : BOOL := FALSE;
    error : BOOL := FALSE;
    status : WORD := 16#0000;
END_VAR

VAR
    buffer : ARRAY[1..100] OF LREAL;
    index : INT := 1;
    count : INT := 0;
    sum : LREAL := 0.0;
    prevCyclic : BOOL := FALSE;
    prevTrigger : BOOL := FALSE;
    prevReset : BOOL := FALSE;
END_VAR

// Reset on rising edge
IF reset AND NOT prevReset THEN
    index := 1;
    count := 0;
    sum := 0.0;
    average := 0.0;
    windowSizeReached := FALSE;
    error := FALSE;
    status := 16#0000;
END_IF;

// Validate window size
IF windowSize < 1 OR windowSize > 100 THEN
    error := TRUE;
    status := 16#8200;
    RETURN;
END_IF;

error := FALSE;
status := 16#0000;

// Process cyclic execution on rising edge
IF cyclicExecution AND NOT prevCyclic THEN
    // Add value
    sum := sum + value;
    buffer[index] := value;
    IF count < windowSize THEN
        count := count + 1;
        windowSizeReached := FALSE;
    ELSE
        sum := sum - buffer[index];
    END_IF;
    average := sum / INT_TO_LREAL(count);
    index := (index MOD windowSize) + 1;
END_IF;

// Process trigger on rising edge (only when cyclicExecution is FALSE)
IF (NOT cyclicExecution) AND trigger AND NOT prevTrigger THEN
    // Add value
    sum := sum + value;
    buffer[index] := value;
    IF count < windowSize THEN
        count := count + 1;
        windowSizeReached := FALSE;
    ELSE
        sum := sum - buffer[index];
    END_IF;
    average := sum / INT_TO_LREAL(count);
    index := (index MOD windowSize) + 1;
END_IF;

// Update previous states
prevCyclic := cyclicExecution;
prevTrigger := trigger;
prevReset := reset;
END_FUNCTION_BLOCK

(* ---- public-medium-03.candidate_02.st ---- *)
FUNCTION_BLOCK FB_MovingAverage
VAR_INPUT
    cyclicExecution : BOOL;
    trigger : BOOL;
    value : LREAL;
    windowSize : INT;
    reset : BOOL;
END_VAR

VAR_OUTPUT
    average : LREAL := 0.0;
    windowSizeReached : BOOL := FALSE;
    error : BOOL := FALSE;
    status : WORD := 16#0000;
END_VAR

VAR
    buffer : ARRAY[1..100] OF LREAL;
    index : INT := 1;
    count : INT := 0;
    sum : LREAL := 0.0;
    prevTrigger : BOOL := FALSE;
END_VAR

// Reset
IF reset THEN
    index := 1;
    count := 0;
    sum := 0.0;
    average := 0.0;
    windowSizeReached := FALSE;
    error := FALSE;
    status := 16#0000;
    RETURN;
END_IF;

// Validate window size
IF windowSize < 1 OR windowSize > 100 THEN
    error := TRUE;
    status := 16#8200;
    RETURN;
END_IF;

error := FALSE;
status := 16#0000;

// Process: cyclic every cycle, or trigger on rising edge
IF cyclicExecution OR (trigger AND NOT prevTrigger) THEN
    sum := sum + value;
    buffer[index] := value;
    IF count < windowSize THEN
        count := count + 1;
        windowSizeReached := FALSE;
    ELSE
        sum := sum - buffer[index];
        windowSizeReached := TRUE;
    END_IF;
    average := sum / INT_TO_LREAL(count);
    index := (index MOD windowSize) + 1;
END_IF;

prevTrigger := trigger;
END_FUNCTION_BLOCK

(* ---- public-medium-03.raw_candidate_01.st ---- *)
FUNCTION_BLOCK FB_MovingAverage
VAR_INPUT
    cyclicExecution : BOOL;
    trigger : BOOL;
    value : LREAL;
    windowSize : INT;
    reset : BOOL;
END_VAR

VAR_OUTPUT
    average : LREAL := 0.0;
    windowSizeReached : BOOL := FALSE;
    error : BOOL := FALSE;
    status : WORD := 16#0000;
END_VAR

VAR
    buffer : ARRAY[1..100] OF LREAL;
    index : INT := 1;
    count : INT := 0;
    sum : LREAL := 0.0;
    prevCyclic : BOOL := FALSE;
    prevTrigger : BOOL := FALSE;
    prevReset : BOOL := FALSE;
END_VAR

// Reset on rising edge
IF reset AND NOT prevReset THEN
    index := 1;
    count := 0;
    sum := 0.0;
    average := 0.0;
    windowSizeReached := FALSE;
    error := FALSE;
    status := 16#0000;
END_IF;

// Validate window size
IF windowSize < 1 OR windowSize > 100 THEN
    error := TRUE;
    status := 16#8200;
    RETURN;
END_IF;

error := FALSE;
status := 16#0000;

// Process cyclic execution on rising edge
IF cyclicExecution AND NOT prevCyclic THEN
    // Add value
    sum := sum + value;
    buffer[index] := value;
    IF count < windowSize THEN
        count := count + 1;
        windowSizeReached := FALSE;
    ELSE
        sum := sum - buffer[index];
    END_IF;
    average := sum / INT_TO_LREAL(count);
    index := (index MOD windowSize) + 1;
END_IF;

// Process trigger on rising edge (only when cyclicExecution is FALSE)
IF (NOT cyclicExecution) AND trigger AND NOT prevTrigger THEN
    // Add value
    sum := sum + value;
    buffer[index] := value;
    IF count < windowSize THEN
        count := count + 1;
        windowSizeReached := FALSE;
    ELSE
        sum := sum - buffer[index];
    END_IF;
    average := sum / INT_TO_LREAL(count);
    index := (index MOD windowSize) + 1;
END_IF;

// Update previous states
prevCyclic := cyclicExecution;
prevTrigger := trigger;
prevReset := reset;
END_FUNCTION_BLOCK

(* ---- public-medium-03.raw_candidate_02.st ---- *)
FUNCTION_BLOCK FB_MovingAverage
VAR_INPUT
    cyclicExecution : BOOL;
    trigger : BOOL;
    value : LREAL;
    windowSize : INT;
    reset : BOOL;
END_VAR

VAR_OUTPUT
    average : LREAL := 0.0;
    windowSizeReached : BOOL := FALSE;
    error : BOOL := FALSE;
    status : WORD := 16#0000;
END_VAR

VAR
    buffer : ARRAY[1..100] OF LREAL;
    index : INT := 1;
    count : INT := 0;
    sum : LREAL := 0.0;
    prevTrigger : BOOL := FALSE;
END_VAR

// Reset
IF reset THEN
    index := 1;
    count := 0;
    sum := 0.0;
    average := 0.0;
    windowSizeReached := FALSE;
    error := FALSE;
    status := 16#0000;
    RETURN;
END_IF;

// Validate window size
IF windowSize < 1 OR windowSize > 100 THEN
    error := TRUE;
    status := 16#8200;
    RETURN;
END_IF;

error := FALSE;
status := 16#0000;

// Process: cyclic every cycle, or trigger on rising edge
IF cyclicExecution OR (trigger AND NOT prevTrigger) THEN
    sum := sum + value;
    buffer[index] := value;
    IF count < windowSize THEN
        count := count + 1;
        windowSizeReached := FALSE;
    ELSE
        sum := sum - buffer[index];
        windowSizeReached := TRUE;
    END_IF;
    average := sum / INT_TO_LREAL(count);
    index := (index MOD windowSize) + 1;
END_IF;

prevTrigger := trigger;
END_FUNCTION_BLOCK

(* ---- public-medium-04.candidate_01.st ---- *)
FUNCTION_BLOCK FB_TemperatureControl
VAR_INPUT
    TemperatureSensorInput : REAL;
    SetTemperature : REAL;
END_VAR

VAR_OUTPUT
    CurrentTemperature : REAL;
    SetTempDisplay : REAL;
    HeaterStatus : BOOL;
    OverheatProtection : BOOL;
    HeaterOutput : BOOL;
END_VAR

VAR
    OverheatTimer : TON;
    CooldownTimer : TON;
    CooldownDone : BOOL;
    HeaterOn : BOOL;
END_VAR

// Update displays
CurrentTemperature := TemperatureSensorInput;
SetTempDisplay := SetTemperature;

// Sensor fault check
IF TemperatureSensorInput < 0.0 OR TemperatureSensorInput > 100.0 THEN
    OverheatProtection := TRUE;
    HeaterOutput := FALSE;
    CooldownTimer(IN := FALSE);
    OverheatTimer(IN := FALSE);
    HeaterStatus := FALSE;
    RETURN;
END_IF;

// Overheat protection cooldown
IF OverheatProtection THEN
    CooldownTimer(IN := TRUE, PT := T#3S);
    CooldownDone := CooldownTimer.Q;
    IF CooldownDone THEN
        OverheatProtection := FALSE;
        CooldownTimer(IN := FALSE);
        HeaterOn := FALSE;
    END_IF;
    HeaterOutput := FALSE;
    HeaterStatus := FALSE;
    RETURN;
END_IF;

// Temperature comparison and heater control
IF TemperatureSensorInput < SetTemperature THEN
    HeaterOn := TRUE;
    OverheatTimer(IN := TRUE, PT := T#5S);
    IF OverheatTimer.Q THEN
        OverheatProtection := TRUE;
        HeaterOn := FALSE;
        HeaterOutput := FALSE;
        OverheatTimer(IN := FALSE);
        RETURN;
    END_IF;
    HeaterOutput := TRUE;
ELSE
    HeaterOn := FALSE;
    HeaterOutput := FALSE;
    OverheatTimer(IN := FALSE);
END_IF;

HeaterStatus := HeaterOutput;

END_FUNCTION_BLOCK

(* ---- public-medium-04.candidate_02.st ---- *)
FUNCTION_BLOCK FB_TemperatureControl
VAR_INPUT
    TemperatureSensorInput : REAL;
    SetTemperature : REAL;
END_VAR

VAR_OUTPUT
    CurrentTemperature : REAL;
    SetTempDisplay : REAL;
    HeaterStatus : BOOL;
    OverheatProtection : BOOL;
    HeaterOutput : BOOL;
END_VAR

VAR
    OverheatTimer : TON;
    CooldownTimer : TON;
    CooldownDone : BOOL;
    HeaterOn : BOOL;
END_VAR

CurrentTemperature := TemperatureSensorInput;
SetTempDisplay := SetTemperature;

IF TemperatureSensorInput < 0.0 OR TemperatureSensorInput > 100.0 THEN
    OverheatProtection := TRUE;
    HeaterOutput := FALSE;
    HeaterStatus := FALSE;
    CooldownTimer(IN := FALSE);
    OverheatTimer(IN := FALSE);
    CooldownDone := FALSE;
    HeaterOn := FALSE;
ELSIF OverheatProtection THEN
    CooldownTimer(IN := TRUE, PT := T#3S);
    CooldownDone := CooldownTimer.Q;
    IF CooldownTimer.Q THEN
        OverheatProtection := FALSE;
        CooldownTimer(IN := FALSE);
        CooldownDone := FALSE;
        HeaterOn := FALSE;
    END_IF;
    HeaterOutput := FALSE;
    HeaterStatus := FALSE;
ELSIF TemperatureSensorInput < SetTemperature THEN
    HeaterOn := TRUE;
    OverheatTimer(IN := TRUE, PT := T#5S);
    IF OverheatTimer.Q THEN
        OverheatProtection := TRUE;
        HeaterOutput := FALSE;
        HeaterStatus := FALSE;
        OverheatTimer(IN := FALSE);
    ELSE
        HeaterOutput := TRUE;
        HeaterStatus := TRUE;
    END_IF;
ELSE
    HeaterOn := FALSE;
    HeaterOutput := FALSE;
    OverheatTimer(IN := FALSE);
    HeaterStatus := FALSE;
END_IF;

END_FUNCTION_BLOCK

(* ---- public-medium-04.raw_candidate_01.st ---- *)
FUNCTION_BLOCK FB_TemperatureControl
VAR_INPUT
    TemperatureSensorInput : REAL;
    SetTemperature : REAL;
END_VAR

VAR_OUTPUT
    CurrentTemperature : REAL;
    SetTempDisplay : REAL;
    HeaterStatus : BOOL;
    OverheatProtection : BOOL;
    HeaterOutput : BOOL;
END_VAR

VAR
    OverheatTimer : TON;
    CooldownTimer : TON;
    CooldownDone : BOOL;
    HeaterOn : BOOL;
END_VAR

// Update displays
CurrentTemperature := TemperatureSensorInput;
SetTempDisplay := SetTemperature;

// Sensor fault check
IF TemperatureSensorInput < 0.0 OR TemperatureSensorInput > 100.0 THEN
    OverheatProtection := TRUE;
    HeaterOutput := FALSE;
    CooldownTimer(IN := FALSE);
    OverheatTimer(IN := FALSE);
    HeaterStatus := FALSE;
    RETURN;
END_IF;

// Overheat protection cooldown
IF OverheatProtection THEN
    CooldownTimer(IN := TRUE, PT := T#3S);
    CooldownDone := CooldownTimer.Q;
    IF CooldownDone THEN
        OverheatProtection := FALSE;
        CooldownTimer(IN := FALSE);
        HeaterOn := FALSE;
    END_IF;
    HeaterOutput := FALSE;
    HeaterStatus := FALSE;
    RETURN;
END_IF;

// Temperature comparison and heater control
IF TemperatureSensorInput < SetTemperature THEN
    HeaterOn := TRUE;
    OverheatTimer(IN := TRUE, PT := T#5S);
    IF OverheatTimer.Q THEN
        OverheatProtection := TRUE;
        HeaterOn := FALSE;
        HeaterOutput := FALSE;
        OverheatTimer(IN := FALSE);
        RETURN;
    END_IF;
    HeaterOutput := TRUE;
ELSE
    HeaterOn := FALSE;
    HeaterOutput := FALSE;
    OverheatTimer(IN := FALSE);
END_IF;

HeaterStatus := HeaterOutput;

END_FUNCTION_BLOCK

(* ---- public-medium-04.raw_candidate_02.st ---- *)
FUNCTION_BLOCK FB_TemperatureControl
VAR_INPUT
    TemperatureSensorInput : REAL;
    SetTemperature : REAL;
END_VAR

VAR_OUTPUT
    CurrentTemperature : REAL;
    SetTempDisplay : REAL;
    HeaterStatus : BOOL;
    OverheatProtection : BOOL;
    HeaterOutput : BOOL;
END_VAR

VAR
    OverheatTimer : TON;
    CooldownTimer : TON;
    CooldownDone : BOOL;
    HeaterOn : BOOL;
END_VAR

CurrentTemperature := TemperatureSensorInput;
SetTempDisplay := SetTemperature;

IF TemperatureSensorInput < 0.0 OR TemperatureSensorInput > 100.0 THEN
    OverheatProtection := TRUE;
    HeaterOutput := FALSE;
    HeaterStatus := FALSE;
    CooldownTimer(IN := FALSE);
    OverheatTimer(IN := FALSE);
    CooldownDone := FALSE;
    HeaterOn := FALSE;
ELSIF OverheatProtection THEN
    CooldownTimer(IN := TRUE, PT := T#3S);
    CooldownDone := CooldownTimer.Q;
    IF CooldownTimer.Q THEN
        OverheatProtection := FALSE;
        CooldownTimer(IN := FALSE);
        CooldownDone := FALSE;
        HeaterOn := FALSE;
    END_IF;
    HeaterOutput := FALSE;
    HeaterStatus := FALSE;
ELSIF TemperatureSensorInput < SetTemperature THEN
    HeaterOn := TRUE;
    OverheatTimer(IN := TRUE, PT := T#5S);
    IF OverheatTimer.Q THEN
        OverheatProtection := TRUE;
        HeaterOutput := FALSE;
        HeaterStatus := FALSE;
        OverheatTimer(IN := FALSE);
    ELSE
        HeaterOutput := TRUE;
        HeaterStatus := TRUE;
    END_IF;
ELSE
    HeaterOn := FALSE;
    HeaterOutput := FALSE;
    OverheatTimer(IN := FALSE);
    HeaterStatus := FALSE;
END_IF;

END_FUNCTION_BLOCK

(* ---- public-medium-05.candidate_01.st ---- *)
FUNCTION_BLOCK ProductionLineControl
VAR_INPUT
    Mode : BOOL;
    ForwardButton : BOOL;
    ReverseButton : BOOL;
    SensorA : BOOL;
    SensorB : BOOL;
    SensorC : BOOL;
    ButtonA : BOOL;
    ButtonB : BOOL;
    ButtonC : BOOL;
END_VAR

VAR_OUTPUT
    MotorForward : BOOL;
    MotorReverse : BOOL;
    CompletionLight : BOOL;
END_VAR

VAR
    State : INT := 0;
    PrevButtonA : BOOL := FALSE;
    PrevButtonB : BOOL := FALSE;
    PrevButtonC : BOOL := FALSE;
END_VAR

IF Mode = FALSE THEN
    MotorForward := ForwardButton AND NOT ReverseButton;
    MotorReverse := ReverseButton AND NOT ForwardButton;
ELSE
    MotorForward := FALSE;
    MotorReverse := FALSE;

    CASE State OF
        0:
            IF SensorA THEN
                State := 1;
            END_IF;

        1:
            IF ButtonA AND NOT PrevButtonA THEN
                MotorForward := TRUE;
                State := 2;
            END_IF;

        2:
            IF SensorB THEN
                MotorForward := FALSE;
                State := 3;
            END_IF;

        3:
            IF ButtonB AND NOT PrevButtonB THEN
                MotorForward := TRUE;
                State := 4;
            END_IF;

        4:
            IF SensorC THEN
                MotorForward := FALSE;
                State := 5;
            END_IF;

        5:
            IF ButtonC AND NOT PrevButtonC THEN
                CompletionLight := TRUE;
                State := 6;
            END_IF;

        6:
            IF NOT SensorC THEN
                CompletionLight := FALSE;
                State := 0;
            END_IF;
    END_CASE;

    PrevButtonA := ButtonA;
    PrevButtonB := ButtonB;
    PrevButtonC := ButtonC;
END_IF;

END_FUNCTION_BLOCK

(* ---- public-medium-05.candidate_02.st ---- *)
FUNCTION_BLOCK ProductionLineControl
VAR_INPUT
    Mode : BOOL;
    ForwardButton : BOOL;
    ReverseButton : BOOL;
    SensorA : BOOL;
    SensorB : BOOL;
    SensorC : BOOL;
    ButtonA : BOOL;
    ButtonB : BOOL;
    ButtonC : BOOL;
END_VAR

VAR_OUTPUT
    MotorForward : BOOL := FALSE;
    MotorReverse : BOOL := FALSE;
    CompletionLight : BOOL := FALSE;
END_VAR

VAR
    State : INT := 0;
    PrevButtonA : BOOL := FALSE;
    PrevButtonB : BOOL := FALSE;
    PrevButtonC : BOOL := FALSE;
END_VAR

IF Mode = FALSE THEN
    MotorForward := ForwardButton AND NOT ReverseButton;
    MotorReverse := ReverseButton AND NOT ForwardButton;
ELSE
    MotorForward := FALSE;
    MotorReverse := FALSE;

    CASE State OF
        0:
            IF SensorA THEN
                State := 1;
            END_IF;

        1:
            IF ButtonA AND NOT PrevButtonA THEN
                MotorForward := TRUE;
                State := 2;
            END_IF;

        2:
            IF SensorB THEN
                MotorForward := FALSE;
                State := 3;
            END_IF;

        3:
            IF ButtonB AND NOT PrevButtonB THEN
                MotorForward := TRUE;
                State := 4;
            END_IF;

        4:
            IF SensorC THEN
                MotorForward := FALSE;
                State := 5;
            END_IF;

        5:
            IF ButtonC AND NOT PrevButtonC THEN
                CompletionLight := TRUE;
                State := 6;
            END_IF;

        6:
            IF NOT SensorC THEN
                CompletionLight := FALSE;
                State := 0;
            END_IF;
    END_CASE;

    PrevButtonA := ButtonA;
    PrevButtonB := ButtonB;
    PrevButtonC := ButtonC;
END_IF;

END_FUNCTION_BLOCK

(* ---- public-medium-05.raw_candidate_01.st ---- *)
FUNCTION_BLOCK ProductionLineControl
VAR_INPUT
    Mode : BOOL;
    ForwardButton : BOOL;
    ReverseButton : BOOL;
    SensorA : BOOL;
    SensorB : BOOL;
    SensorC : BOOL;
    ButtonA : BOOL;
    ButtonB : BOOL;
    ButtonC : BOOL;
END_VAR

VAR_OUTPUT
    MotorForward : BOOL;
    MotorReverse : BOOL;
    CompletionLight : BOOL;
END_VAR

VAR
    State : INT := 0;
    PrevButtonA : BOOL := FALSE;
    PrevButtonB : BOOL := FALSE;
    PrevButtonC : BOOL := FALSE;
END_VAR

IF Mode = FALSE THEN
    MotorForward := ForwardButton AND NOT ReverseButton;
    MotorReverse := ReverseButton AND NOT ForwardButton;
ELSE
    MotorForward := FALSE;
    MotorReverse := FALSE;

    CASE State OF
        0:
            IF SensorA THEN
                State := 1;
            END_IF

        1:
            IF ButtonA AND NOT PrevButtonA THEN
                MotorForward := TRUE;
                State := 2;
            END_IF

        2:
            IF SensorB THEN
                MotorForward := FALSE;
                State := 3;
            END_IF

        3:
            IF ButtonB AND NOT PrevButtonB THEN
                MotorForward := TRUE;
                State := 4;
            END_IF

        4:
            IF SensorC THEN
                MotorForward := FALSE;
                State := 5;
            END_IF

        5:
            IF ButtonC AND NOT PrevButtonC THEN
                CompletionLight := TRUE;
                State := 6;
            END_IF

        6:
            IF NOT SensorC THEN
                CompletionLight := FALSE;
                State := 0;
            END_IF
    END_CASE;

    PrevButtonA := ButtonA;
    PrevButtonB := ButtonB;
    PrevButtonC := ButtonC;
END_IF

END_FUNCTION_BLOCK

(* ---- public-medium-05.raw_candidate_02.st ---- *)
FUNCTION_BLOCK ProductionLineControl
VAR_INPUT
    Mode : BOOL;
    ForwardButton : BOOL;
    ReverseButton : BOOL;
    SensorA : BOOL;
    SensorB : BOOL;
    SensorC : BOOL;
    ButtonA : BOOL;
    ButtonB : BOOL;
    ButtonC : BOOL;
END_VAR

VAR_OUTPUT
    MotorForward : BOOL := FALSE;
    MotorReverse : BOOL := FALSE;
    CompletionLight : BOOL := FALSE;
END_VAR

VAR
    State : INT := 0;
    PrevButtonA : BOOL := FALSE;
    PrevButtonB : BOOL := FALSE;
    PrevButtonC : BOOL := FALSE;
END_VAR

IF Mode = FALSE THEN
    MotorForward := ForwardButton AND NOT ReverseButton;
    MotorReverse := ReverseButton AND NOT ForwardButton;
ELSE
    MotorForward := FALSE;
    MotorReverse := FALSE;

    CASE State OF
        0:
            IF SensorA THEN
                State := 1;
            END_IF;

        1:
            IF ButtonA AND NOT PrevButtonA THEN
                MotorForward := TRUE;
                State := 2;
            END_IF;

        2:
            IF SensorB THEN
                MotorForward := FALSE;
                State := 3;
            END_IF;

        3:
            IF ButtonB AND NOT PrevButtonB THEN
                MotorForward := TRUE;
                State := 4;
            END_IF;

        4:
            IF SensorC THEN
                MotorForward := FALSE;
                State := 5;
            END_IF;

        5:
            IF ButtonC AND NOT PrevButtonC THEN
                CompletionLight := TRUE;
                State := 6;
            END_IF;

        6:
            IF NOT SensorC THEN
                CompletionLight := FALSE;
                State := 0;
            END_IF;
    END_CASE;

    PrevButtonA := ButtonA;
    PrevButtonB := ButtonB;
    PrevButtonC := ButtonC;
END_IF;

END_FUNCTION_BLOCK

(* ---- public-medium-06.candidate_01.st ---- *)
FUNCTION_BLOCK SlabThicknessAlarm
VAR_INPUT
    THICKNESS_FAULT : BOOL;
    THICKNESS_SIGNAL_VALID : BOOL;
    CUTTING_RUN : BOOL;
    FaultTimestamp : DINT;
    CycleTime : TIME;
END_VAR

VAR_OUTPUT
    THICKNESS_ALARM : BOOL;
    Slab_Fault_Counter : UINT;
    Slab_Runtime_Accumulator : LTIME;
    Slab_Fault_History : ARRAY[0..4] OF DINT;
END_VAR

VAR
    AlarmHoldTimer : TON;
    FallEdgeFault : R_TRIG;
    PreviousFaultValid : BOOL := FALSE;
    PreviousSignalValid : BOOL := FALSE;
END_VAR

// Detect FALSE-to-TRUE transition of valid fault signal
IF THICKNESS_SIGNAL_VALID AND THICKNESS_FAULT AND NOT PreviousFaultValid THEN
    // Shift history and record new fault
    Slab_Fault_History[4] := Slab_Fault_History[3];
    Slab_Fault_History[3] := Slab_Fault_History[2];
    Slab_Fault_History[2] := Slab_Fault_History[1];
    Slab_Fault_History[1] := Slab_Fault_History[0];
    Slab_Fault_History[0] := FaultTimestamp;
    Slab_Fault_Counter := Slab_Fault_Counter + 1;
END_IF;

// Alarm control
IF NOT THICKNESS_SIGNAL_VALID THEN
    THICKNESS_ALARM := FALSE;
    AlarmHoldTimer(IN := FALSE);
ELSE
    IF THICKNESS_FAULT THEN
        THICKNESS_ALARM := TRUE;
        AlarmHoldTimer(IN := FALSE);
    ELSE
        FallEdgeFault(CLK := PreviousFaultValid AND NOT THICKNESS_FAULT);
        IF FallEdgeFault.Q THEN
            AlarmHoldTimer(IN := TRUE, PT := T#500ms);
        END_IF;
        IF AlarmHoldTimer.Q THEN
            THICKNESS_ALARM := FALSE;
        END_IF;
    END_IF;
END_IF;

// Runtime accumulation
IF NOT THICKNESS_SIGNAL_VALID THEN
    Slab_Runtime_Accumulator := LTIME#0s;
ELSE
    IF CUTTING_RUN AND NOT THICKNESS_FAULT THEN
        Slab_Runtime_Accumulator := Slab_Runtime_Accumulator + LTIME_TO_LINT(CycleTime);
    END_IF;
END_IF;

// Update state tracking
PreviousFaultValid := THICKNESS_FAULT;
PreviousSignalValid := THICKNESS_SIGNAL_VALID;

END_FUNCTION_BLOCK

(* ---- public-medium-06.candidate_02.st ---- *)
FUNCTION_BLOCK SlabThicknessAlarm
VAR_INPUT
    THICKNESS_FAULT : BOOL;
    THICKNESS_SIGNAL_VALID : BOOL;
    CUTTING_RUN : BOOL;
    FaultTimestamp : DINT;
    CycleTime : TIME;
END_VAR

VAR_OUTPUT
    THICKNESS_ALARM : BOOL;
    Slab_Fault_Counter : UINT;
    Slab_Runtime_Accumulator : LTIME;
    Slab_Fault_History : ARRAY[0..4] OF DINT;
END_VAR

VAR
    AlarmHoldTimer : TON;
    FallEdgeFault : R_TRIG;
    PreviousFaultValid : BOOL := FALSE;
    PreviousSignalValid : BOOL := FALSE;
END_VAR

// Detect FALSE-to-TRUE transition of valid fault signal
IF THICKNESS_SIGNAL_VALID AND THICKNESS_FAULT AND NOT PreviousFaultValid THEN
    Slab_Fault_History[4] := Slab_Fault_History[3];
    Slab_Fault_History[3] := Slab_Fault_History[2];
    Slab_Fault_History[2] := Slab_Fault_History[1];
    Slab_Fault_History[1] := Slab_Fault_History[0];
    Slab_Fault_History[0] := FaultTimestamp;
    Slab_Fault_Counter := Slab_Fault_Counter + 1;
END_IF;

// Alarm control
IF NOT THICKNESS_SIGNAL_VALID THEN
    THICKNESS_ALARM := FALSE;
    AlarmHoldTimer(IN := FALSE);
ELSE
    IF THICKNESS_FAULT THEN
        THICKNESS_ALARM := TRUE;
        AlarmHoldTimer(IN := FALSE);
    ELSE
        FallEdgeFault(CLK := PreviousFaultValid AND NOT THICKNESS_FAULT);
        IF FallEdgeFault.Q THEN
            AlarmHoldTimer(IN := TRUE, PT := T#500ms);
        END_IF;
        IF AlarmHoldTimer.Q THEN
            THICKNESS_ALARM := FALSE;
        END_IF;
    END_IF;
END_IF;

// Runtime accumulation
IF CUTTING_RUN AND THICKNESS_SIGNAL_VALID AND NOT THICKNESS_FAULT THEN
    Slab_Runtime_Accumulator := Slab_Runtime_Accumulator + TIME_TO_LTIME(CycleTime);
END_IF;

// Update state tracking
PreviousFaultValid := THICKNESS_FAULT;
PreviousSignalValid := THICKNESS_SIGNAL_VALID;

END_FUNCTION_BLOCK

(* ---- public-medium-06.raw_candidate_01.st ---- *)
FUNCTION_BLOCK SlabThicknessAlarm
VAR_INPUT
    THICKNESS_FAULT : BOOL;
    THICKNESS_SIGNAL_VALID : BOOL;
    CUTTING_RUN : BOOL;
    FaultTimestamp : DINT;
    CycleTime : TIME;
END_VAR

VAR_OUTPUT
    THICKNESS_ALARM : BOOL;
    Slab_Fault_Counter : UINT;
    Slab_Runtime_Accumulator : LTIME;
    Slab_Fault_History : ARRAY[0..4] OF DINT;
END_VAR

VAR
    AlarmHoldTimer : TON;
    FallEdgeFault : R_TRIG;
    PreviousFaultValid : BOOL := FALSE;
    PreviousSignalValid : BOOL := FALSE;
END_VAR

// Detect FALSE-to-TRUE transition of valid fault signal
IF THICKNESS_SIGNAL_VALID AND THICKNESS_FAULT AND NOT PreviousFaultValid THEN
    // Shift history and record new fault
    Slab_Fault_History[4] := Slab_Fault_History[3];
    Slab_Fault_History[3] := Slab_Fault_History[2];
    Slab_Fault_History[2] := Slab_Fault_History[1];
    Slab_Fault_History[1] := Slab_Fault_History[0];
    Slab_Fault_History[0] := FaultTimestamp;
    Slab_Fault_Counter := Slab_Fault_Counter + 1;
END_IF;

// Alarm control
IF NOT THICKNESS_SIGNAL_VALID THEN
    THICKNESS_ALARM := FALSE;
    AlarmHoldTimer(IN := FALSE);
ELSE
    IF THICKNESS_FAULT THEN
        THICKNESS_ALARM := TRUE;
        AlarmHoldTimer(IN := FALSE);
    ELSE
        FallEdgeFault(CLK := PreviousFaultValid AND NOT THICKNESS_FAULT);
        IF FallEdgeFault.Q THEN
            AlarmHoldTimer(IN := TRUE, PT := T#500ms);
        END_IF;
        IF AlarmHoldTimer.Q THEN
            THICKNESS_ALARM := FALSE;
        END_IF;
    END_IF;
END_IF;

// Runtime accumulation
IF NOT THICKNESS_SIGNAL_VALID THEN
    Slab_Runtime_Accumulator := LTIME#0s;
ELSE
    IF CUTTING_RUN AND NOT THICKNESS_FAULT THEN
        Slab_Runtime_Accumulator := Slab_Runtime_Accumulator + LTIME_TO_LINT(CycleTime);
    END_IF;
END_IF;

// Update state tracking
PreviousFaultValid := THICKNESS_FAULT;
PreviousSignalValid := THICKNESS_SIGNAL_VALID;

END_FUNCTION_BLOCK

(* ---- public-medium-06.raw_candidate_02.st ---- *)
FUNCTION_BLOCK SlabThicknessAlarm
VAR_INPUT
    THICKNESS_FAULT : BOOL;
    THICKNESS_SIGNAL_VALID : BOOL;
    CUTTING_RUN : BOOL;
    FaultTimestamp : DINT;
    CycleTime : TIME;
END_VAR

VAR_OUTPUT
    THICKNESS_ALARM : BOOL;
    Slab_Fault_Counter : UINT;
    Slab_Runtime_Accumulator : LTIME;
    Slab_Fault_History : ARRAY[0..4] OF DINT;
END_VAR

VAR
    AlarmHoldTimer : TON;
    FallEdgeFault : R_TRIG;
    PreviousFaultValid : BOOL := FALSE;
    PreviousSignalValid : BOOL := FALSE;
END_VAR

// Detect FALSE-to-TRUE transition of valid fault signal
IF THICKNESS_SIGNAL_VALID AND THICKNESS_FAULT AND NOT PreviousFaultValid THEN
    Slab_Fault_History[4] := Slab_Fault_History[3];
    Slab_Fault_History[3] := Slab_Fault_History[2];
    Slab_Fault_History[2] := Slab_Fault_History[1];
    Slab_Fault_History[1] := Slab_Fault_History[0];
    Slab_Fault_History[0] := FaultTimestamp;
    Slab_Fault_Counter := Slab_Fault_Counter + 1;
END_IF;

// Alarm control
IF NOT THICKNESS_SIGNAL_VALID THEN
    THICKNESS_ALARM := FALSE;
    AlarmHoldTimer(IN := FALSE);
ELSE
    IF THICKNESS_FAULT THEN
        THICKNESS_ALARM := TRUE;
        AlarmHoldTimer(IN := FALSE);
    ELSE
        FallEdgeFault(CLK := PreviousFaultValid AND NOT THICKNESS_FAULT);
        IF FallEdgeFault.Q THEN
            AlarmHoldTimer(IN := TRUE, PT := T#500ms);
        END_IF;
        IF AlarmHoldTimer.Q THEN
            THICKNESS_ALARM := FALSE;
        END_IF;
    END_IF;
END_IF;

// Runtime accumulation
IF CUTTING_RUN AND THICKNESS_SIGNAL_VALID AND NOT THICKNESS_FAULT THEN
    Slab_Runtime_Accumulator := Slab_Runtime_Accumulator + TIME_TO_LTIME(CycleTime);
END_IF;

// Update state tracking
PreviousFaultValid := THICKNESS_FAULT;
PreviousSignalValid := THICKNESS_SIGNAL_VALID;

END_FUNCTION_BLOCK

(* ---- public-medium-07.candidate_01.st ---- *)
FUNCTION_BLOCK HVAC_Controller
VAR_INPUT
    OCCUPANCY_DETECTED      : BOOL;
    ENERGY_SAVING_MODE      : BOOL;
    HVAC_MODE_SELECTOR      : INT;
END_VAR

VAR_OUTPUT
    SUPPLY_FAN_RUN          : BOOL;
    TEMP_SETPOINT_ADJUST    : INT;
END_VAR

VAR
    OccupancyTimer          : TON;
    OccupancyStartTime      : LTIME;
    FanDelayActive          : BOOL := FALSE;
    FanDelayElapsed         : BOOL := FALSE;
    PreviousOccupancy       : BOOL := FALSE;
END_VAR

// Fan control logic
IF NOT OCCUPANCY_DETECTED OR (HVAC_MODE_SELECTOR = 3) THEN
    // Reset delay when occupancy lost or Night mode selected
    FanDelayActive := FALSE;
    FanDelayElapsed := FALSE;
    SUPPLY_FAN_RUN := FALSE;
    OccupancyTimer(IN := FALSE);
ELSIF OCCUPANCY_DETECTED AND (HVAC_MODE_SELECTOR <> 3) THEN
    // Start delay when occupancy detected and not in Night mode
    IF NOT FanDelayActive THEN
        FanDelayActive := TRUE;
        OccupancyTimer(IN := FALSE);
    END_IF;
    OccupancyTimer(IN := TRUE, PT := T#30S);
    FanDelayElapsed := OccupancyTimer.Q;
    SUPPLY_FAN_RUN := FanDelayElapsed;
ELSE
    // Default to off
    SUPPLY_FAN_RUN := FALSE;
END_IF;

// Temperature setpoint calculation
CASE HVAC_MODE_SELECTOR OF
    0: // Auto mode
        IF OCCUPANCY_DETECTED THEN
            TEMP_SETPOINT_ADJUST := 0;
        ELSE
            IF ENERGY_SAVING_MODE THEN
                TEMP_SETPOINT_ADJUST := 3;
            ELSE
                TEMP_SETPOINT_ADJUST := 2;
            END_IF;
        END_IF;

    1: // Comfort mode
        IF OCCUPANCY_DETECTED THEN
            TEMP_SETPOINT_ADJUST := 0;
        ELSE
            TEMP_SETPOINT_ADJUST := 1;
        END_IF;

    2: // Economy mode
        IF OCCUPANCY_DETECTED THEN
            TEMP_SETPOINT_ADJUST := 0;
        ELSE
            TEMP_SETPOINT_ADJUST := 4;
        END_IF;

    3: // Night mode
        TEMP_SETPOINT_ADJUST := 4;

ELSE
    TEMP_SETPOINT_ADJUST := 0;
END_CASE;

// Clamp to ±4°C
IF TEMP_SETPOINT_ADJUST > 4 THEN
    TEMP_SETPOINT_ADJUST := 4;
ELSIF TEMP_SETPOINT_ADJUST < -4 THEN
    TEMP_SETPOINT_ADJUST := -4;
END_IF;

PreviousOccupancy := OCCUPANCY_DETECTED;

END_FUNCTION_BLOCK

(* ---- public-medium-07.raw_candidate_01.st ---- *)
FUNCTION_BLOCK HVAC_Controller
VAR_INPUT
    OCCUPANCY_DETECTED      : BOOL;
    ENERGY_SAVING_MODE      : BOOL;
    HVAC_MODE_SELECTOR      : INT;
END_VAR

VAR_OUTPUT
    SUPPLY_FAN_RUN          : BOOL;
    TEMP_SETPOINT_ADJUST    : INT;
END_VAR

VAR
    OccupancyTimer          : TON;
    OccupancyStartTime      : LTIME;
    FanDelayActive          : BOOL := FALSE;
    FanDelayElapsed         : BOOL := FALSE;
    PreviousOccupancy       : BOOL := FALSE;
END_VAR

// Fan control logic
IF NOT OCCUPANCY_DETECTED OR (HVAC_MODE_SELECTOR = 3) THEN
    // Reset delay when occupancy lost or Night mode selected
    FanDelayActive := FALSE;
    FanDelayElapsed := FALSE;
    SUPPLY_FAN_RUN := FALSE;
    OccupancyTimer(IN := FALSE);
ELSIF OCCUPANCY_DETECTED AND (HVAC_MODE_SELECTOR <> 3) THEN
    // Start delay when occupancy detected and not in Night mode
    IF NOT FanDelayActive THEN
        FanDelayActive := TRUE;
        OccupancyTimer(IN := FALSE);
    END_IF
    OccupancyTimer(IN := TRUE, PT := T#30S);
    FanDelayElapsed := OccupancyTimer.Q;
    SUPPLY_FAN_RUN := FanDelayElapsed;
ELSE
    // Default to off
    SUPPLY_FAN_RUN := FALSE;
END_IF;

// Temperature setpoint calculation
CASE HVAC_MODE_SELECTOR OF
    0: // Auto mode
        IF OCCUPANCY_DETECTED THEN
            TEMP_SETPOINT_ADJUST := 0;
        ELSE
            IF ENERGY_SAVING_MODE THEN
                TEMP_SETPOINT_ADJUST := 3;
            ELSE
                TEMP_SETPOINT_ADJUST := 2;
            END_IF;
        END_IF;

    1: // Comfort mode
        IF OCCUPANCY_DETECTED THEN
            TEMP_SETPOINT_ADJUST := 0;
        ELSE
            TEMP_SETPOINT_ADJUST := 1;
        END_IF;

    2: // Economy mode
        IF OCCUPANCY_DETECTED THEN
            TEMP_SETPOINT_ADJUST := 0;
        ELSE
            TEMP_SETPOINT_ADJUST := 4;
        END_IF;

    3: // Night mode
        TEMP_SETPOINT_ADJUST := 4;

ELSE
    TEMP_SETPOINT_ADJUST := 0;
END_CASE;

// Clamp to ±4°C
IF TEMP_SETPOINT_ADJUST > 4 THEN
    TEMP_SETPOINT_ADJUST := 4;
ELSIF TEMP_SETPOINT_ADJUST < -4 THEN
    TEMP_SETPOINT_ADJUST := -4;
END_IF;

PreviousOccupancy := OCCUPANCY_DETECTED;

END_FUNCTION_BLOCK

(* ---- public-medium-08.candidate_01.st ---- *)
FUNCTION_BLOCK IPv4Parser
VAR_INPUT
    ipText : STRING(254);
END_VAR
VAR_OUTPUT
    ipValue : UDINT;
END_VAR
VAR
    currentPos : INT;
    segmentLen : INT;
    segmentValue : UDINT;
    dotCount : INT;
    charCode : INT;
    ch : CHAR;
END_VAR

ipValue := 0;

// Basic length validation
IF LEN(ipText) < 7 OR LEN(ipText) > 15 THEN
    RETURN;
END_IF;

currentPos := 1;
dotCount := 0;

WHILE dotCount < 3 AND currentPos <= LEN(ipText) DO
    // Extract one segment
    segmentValue := 0;
    segmentLen := 0;

    WHILE currentPos <= LEN(ipText) DO
        ch := MID(ipText, 1, currentPos);
        charCode := CHAR_TO_INT(ch);

        IF charCode = 46 THEN // '.'
            EXIT;
        ELSIF charCode >= 48 AND charCode <= 57 THEN
            segmentValue := segmentValue * 10 + TO_UDINT(charCode - 48);
            segmentLen := segmentLen + 1;
            currentPos := currentPos + 1;
        ELSE
            ipValue := 0;
            RETURN;
        END_IF;
    END_WHILE;

    // Validate segment
    IF segmentLen = 0 OR segmentLen > 3 THEN
        ipValue := 0;
        RETURN;
    END_IF;

    IF segmentValue > 255 THEN
        ipValue := 0;
        RETURN;
    END_IF;

    // Add to result in network byte order
    ipValue := SHL(ipValue, 8) OR segmentValue;
    dotCount := dotCount + 1;

    // Move to next position after dot
    currentPos := currentPos + 1;
END_WHILE;

// Validate exactly 3 dots (4 segments)
IF dotCount <> 3 THEN
    ipValue := 0;
    RETURN;
END_IF;

// Ensure no content after 4th segment
IF currentPos <= LEN(ipText) THEN
    ipValue := 0;
    RETURN;
END_IF;

END_FUNCTION_BLOCK

(* ---- public-medium-08.candidate_02.st ---- *)
FUNCTION_BLOCK IPv4Parser
VAR_INPUT
    ipText : STRING(254);
END_VAR
VAR_OUTPUT
    ipValue : UDINT;
END_VAR
VAR
    currentPos : INT;
    segmentLen : INT;
    segmentValue : UDINT;
    dotCount : INT;
    ch : STRING(1);
    charVal : INT;
END_VAR

ipValue := 0;

// Basic length validation
IF LEN(ipText) < 7 OR LEN(ipText) > 15 THEN
    RETURN;
END_IF;

currentPos := 1;
dotCount := 0;

WHILE dotCount < 3 AND currentPos <= LEN(ipText) DO
    segmentValue := 0;
    segmentLen := 0;

    WHILE currentPos <= LEN(ipText) DO
        ch := MID(ipText, 1, currentPos);

        IF LEN(ch) = 1 AND MID(ch, 1, 1) = '.' THEN
            EXIT;
        END_IF;

        charVal := INT(MID(ipText, 1, currentPos));

        IF charVal >= 48 AND charVal <= 57 THEN
            segmentValue := segmentValue * 10 + UDINT(DINT(charVal - 48));
            segmentLen := segmentLen + 1;
            currentPos := currentPos + 1;
        ELSE
            ipValue := 0;
            RETURN;
        END_IF;
    END_WHILE;

    IF segmentLen = 0 OR segmentLen > 3 THEN
        ipValue := 0;
        RETURN;
    END_IF;

    IF segmentValue > 255 THEN
        ipValue := 0;
        RETURN;
    END_IF;

    ipValue := SHL(ipValue, 8) OR segmentValue;
    dotCount := dotCount + 1;

    IF currentPos <= LEN(ipText) THEN
        currentPos := currentPos + 1;
    END_IF;
END_WHILE;

IF dotCount <> 3 THEN
    ipValue := 0;
    RETURN;
END_IF;

IF currentPos <= LEN(ipText) AND MID(ipText, 1, currentPos) <> '.' THEN
    ipValue := 0;
    RETURN;
END_IF;

END_FUNCTION_BLOCK

(* ---- public-medium-08.raw_candidate_01.st ---- *)
FUNCTION_BLOCK IPv4Parser
VAR_INPUT
    ipText : STRING(254);
END_VAR
VAR_OUTPUT
    ipValue : UDINT;
END_VAR
VAR
    currentPos : INT;
    segmentLen : INT;
    segmentValue : UDINT;
    dotCount : INT;
    charCode : INT;
    ch : CHAR;
END_VAR

ipValue := 0;

// Basic length validation
IF LEN(ipText) < 7 OR LEN(ipText) > 15 THEN
    RETURN;
END_IF

currentPos := 1;
dotCount := 0;

WHILE dotCount < 3 AND currentPos <= LEN(ipText) DO
    // Extract one segment
    segmentValue := 0;
    segmentLen := 0;

    WHILE currentPos <= LEN(ipText) DO
        ch := MID(ipText, 1, currentPos);
        charCode := CHAR_TO_INT(ch);

        IF charCode = 46 THEN // '.'
            EXIT;
        ELSIF charCode >= 48 AND charCode <= 57 THEN
            segmentValue := segmentValue * 10 + TO_UDINT(charCode - 48);
            segmentLen := segmentLen + 1;
            currentPos := currentPos + 1;
        ELSE
            ipValue := 0;
            RETURN;
        END_IF
    END_WHILE

    // Validate segment
    IF segmentLen = 0 OR segmentLen > 3 THEN
        ipValue := 0;
        RETURN;
    END_IF

    IF segmentValue > 255 THEN
        ipValue := 0;
        RETURN;
    END_IF

    // Add to result in network byte order
    ipValue := SHL(ipValue, 8) OR segmentValue;
    dotCount := dotCount + 1;

    // Move to next position after dot
    currentPos := currentPos + 1;
END_WHILE

// Validate exactly 3 dots (4 segments)
IF dotCount <> 3 THEN
    ipValue := 0;
    RETURN;
END_IF

// Ensure no content after 4th segment
IF currentPos <= LEN(ipText) THEN
    ipValue := 0;
    RETURN;
END_IF

END_FUNCTION_BLOCK

(* ---- public-medium-08.raw_candidate_02.st ---- *)
FUNCTION_BLOCK IPv4Parser
VAR_INPUT
    ipText : STRING(254);
END_VAR
VAR_OUTPUT
    ipValue : UDINT;
END_VAR
VAR
    currentPos : INT;
    segmentLen : INT;
    segmentValue : UDINT;
    dotCount : INT;
    ch : STRING(1);
    charVal : INT;
END_VAR

ipValue := 0;

// Basic length validation
IF LEN(ipText) < 7 OR LEN(ipText) > 15 THEN
    RETURN;
END_IF;

currentPos := 1;
dotCount := 0;

WHILE dotCount < 3 AND currentPos <= LEN(ipText) DO
    segmentValue := 0;
    segmentLen := 0;

    WHILE currentPos <= LEN(ipText) DO
        ch := MID(ipText, 1, currentPos);

        IF LEN(ch) = 1 AND MID(ch, 1, 1) = '.' THEN
            EXIT;
        END_IF;

        charVal := INT(MID(ipText, 1, currentPos));

        IF charVal >= 48 AND charVal <= 57 THEN
            segmentValue := segmentValue * 10 + UDINT(DINT(charVal - 48));
            segmentLen := segmentLen + 1;
            currentPos := currentPos + 1;
        ELSE
            ipValue := 0;
            RETURN;
        END_IF;
    END_WHILE;

    IF segmentLen = 0 OR segmentLen > 3 THEN
        ipValue := 0;
        RETURN;
    END_IF;

    IF segmentValue > 255 THEN
        ipValue := 0;
        RETURN;
    END_IF;

    ipValue := SHL(ipValue, 8) OR segmentValue;
    dotCount := dotCount + 1;

    IF currentPos <= LEN(ipText) THEN
        currentPos := currentPos + 1;
    END_IF;
END_WHILE;

IF dotCount <> 3 THEN
    ipValue := 0;
    RETURN;
END_IF;

IF currentPos <= LEN(ipText) AND MID(ipText, 1, currentPos) <> '.' THEN
    ipValue := 0;
    RETURN;
END_IF;

END_FUNCTION_BLOCK

(* ---- self-easy-01.candidate_01.st ---- *)
FUNCTION_BLOCK FB
VAR
    prevAvgOut : REAL := 0.0;
END_VAR
VAR_INPUT
    enable     : BOOL;
    values     : ARRAY[1..8] OF INT;
    count      : INT;
    avgEnable  : BOOL;
END_VAR
VAR_OUTPUT
    avgOut : REAL;
END_VAR
VAR_TEMP
    sum : DINT;
    effectiveCount : INT;
END_VAR

    // Calculate only when enabled, averaging is active, and we have valid samples
    IF enable AND avgEnable AND count > 0 THEN
        // Clamp count to valid array bounds
        IF count > 8 THEN
            effectiveCount := 8;
        ELSE
            effectiveCount := count;
        END_IF;

        // Accumulate sum in DINT to avoid overflow
        sum := 0;
        IF effectiveCount >= 1 THEN
            sum := sum + values[1];
        END_IF;
        IF effectiveCount >= 2 THEN
            sum := sum + values[2];
        END_IF;
        IF effectiveCount >= 3 THEN
            sum := sum + values[3];
        END_IF;
        IF effectiveCount >= 4 THEN
            sum := sum + values[4];
        END_IF;
        IF effectiveCount >= 5 THEN
            sum := sum + values[5];
        END_IF;
        IF effectiveCount >= 6 THEN
            sum := sum + values[6];
        END_IF;
        IF effectiveCount >= 7 THEN
            sum := sum + values[7];
        END_IF;
        IF effectiveCount >= 8 THEN
            sum := sum + values[8];
        END_IF;

        // Compute average as REAL
        avgOut := DINT_TO_REAL(sum) / DINT_TO_REAL(effectiveCount);
    ELSE
        // Hold previous value when disabled or no valid samples
        avgOut := prevAvgOut;
    END_IF;

    // Update latched output for next scan
    prevAvgOut := avgOut;
END_FUNCTION_BLOCK

(* ---- self-easy-01.raw_candidate_01.st ---- *)
FUNCTION_BLOCK FB
VAR
    prevAvgOut : REAL := 0.0;
END_VAR
VAR_INPUT
    enable     : BOOL;
    values     : ARRAY[1..8] OF INT;
    count      : INT;
    avgEnable  : BOOL;
END_VAR
VAR_OUTPUT
    avgOut : REAL;
END_VAR
VAR_TEMP
    sum : DINT;
    effectiveCount : INT;
END_VAR

    // Calculate only when enabled, averaging is active, and we have valid samples
    IF enable AND avgEnable AND count > 0 THEN
        // Clamp count to valid array bounds
        IF count > 8 THEN
            effectiveCount := 8;
        ELSE
            effectiveCount := count;
        END_IF;

        // Accumulate sum in DINT to avoid overflow
        sum := 0;
        IF effectiveCount >= 1 THEN
            sum := sum + values[1];
        END_IF;
        IF effectiveCount >= 2 THEN
            sum := sum + values[2];
        END_IF;
        IF effectiveCount >= 3 THEN
            sum := sum + values[3];
        END_IF;
        IF effectiveCount >= 4 THEN
            sum := sum + values[4];
        END_IF;
        IF effectiveCount >= 5 THEN
            sum := sum + values[5];
        END_IF;
        IF effectiveCount >= 6 THEN
            sum := sum + values[6];
        END_IF;
        IF effectiveCount >= 7 THEN
            sum := sum + values[7];
        END_IF;
        IF effectiveCount >= 8 THEN
            sum := sum + values[8];
        END_IF;

        // Compute average as REAL
        avgOut := DINT_TO_REAL(sum) / DINT_TO_REAL(effectiveCount);
    ELSE
        // Hold previous value when disabled or no valid samples
        avgOut := prevAvgOut;
    END_IF;

    // Update latched output for next scan
    prevAvgOut := avgOut;
END_FUNCTION_BLOCK

(* ---- self-easy-02.candidate_01.st ---- *)
FUNCTION_BLOCK FB
VAR_INPUT
    tankLevel   : REAL;
    outletFlow  : REAL;
    inletPermit : BOOL;
    resetBtn    : BOOL;
END_VAR
VAR_OUTPUT
    pumpRun        : BOOL;
    alarmHigh      : BOOL;
    alarmLow       : BOOL;
    outletValveOpen: BOOL;
END_VAR
VAR
    prevResetBtn : BOOL := FALSE;
    prevAlarmHigh: BOOL := FALSE;
    prevAlarmLow : BOOL := FALSE;
END_VAR
VAR
    resetRising : BOOL;
END_VAR

resetRising := resetBtn AND NOT prevResetBtn;

IF tankLevel >= 85.0 THEN
    alarmHigh := TRUE;
ELSIF resetRising AND NOT (tankLevel >= 85.0) THEN
    alarmHigh := FALSE;
ELSE
    alarmHigh := prevAlarmHigh;
END_IF;

IF tankLevel <= 15.0 THEN
    alarmLow := TRUE;
ELSIF resetRising AND NOT (tankLevel <= 15.0) THEN
    alarmLow := FALSE;
ELSE
    alarmLow := prevAlarmLow;
END_IF;

pumpRun := (NOT alarmHigh) AND (NOT alarmLow) AND inletPermit;

outletValveOpen := NOT alarmLow;

prevResetBtn  := resetBtn;
prevAlarmHigh := alarmHigh;
prevAlarmLow  := alarmLow;
END_FUNCTION_BLOCK

(* ---- self-easy-02.raw_candidate_01.st ---- *)
FUNCTION_BLOCK FB
VAR_INPUT
    tankLevel   : REAL;
    outletFlow  : REAL;
    inletPermit : BOOL;
    resetBtn    : BOOL;
END_VAR
VAR_OUTPUT
    pumpRun        : BOOL;
    alarmHigh      : BOOL;
    alarmLow       : BOOL;
    outletValveOpen: BOOL;
END_VAR
VAR
    prevResetBtn : BOOL := FALSE;
    prevAlarmHigh: BOOL := FALSE;
    prevAlarmLow : BOOL := FALSE;
END_VAR
VAR
    resetRising : BOOL;
END_VAR

resetRising := resetBtn AND NOT prevResetBtn;

IF tankLevel >= 85.0 THEN
    alarmHigh := TRUE;
ELSIF resetRising AND NOT (tankLevel >= 85.0) THEN
    alarmHigh := FALSE;
ELSE
    alarmHigh := prevAlarmHigh;
END_IF;

IF tankLevel <= 15.0 THEN
    alarmLow := TRUE;
ELSIF resetRising AND NOT (tankLevel <= 15.0) THEN
    alarmLow := FALSE;
ELSE
    alarmLow := prevAlarmLow;
END_IF;

pumpRun := (NOT alarmHigh) AND (NOT alarmLow) AND inletPermit;

outletValveOpen := NOT alarmLow;

prevResetBtn  := resetBtn;
prevAlarmHigh := alarmHigh;
prevAlarmLow  := alarmLow;
END_FUNCTION_BLOCK

(* ---- self-hard-01.candidate_01.st ---- *)
FUNCTION_BLOCK FB
VAR_INPUT
    flowLow   : BOOL;
    ackBtn    : BOOL;
    sensorOK  : BOOL;
END_VAR
VAR_OUTPUT
    alarmActive : BOOL;
    alarmAcked  : BOOL;
    highHigh    : BOOL;
END_VAR
VAR
    prev_flowLow   : BOOL := FALSE;
    prev_ackBtn    : BOOL := FALSE;
    prev_alarmAcked : BOOL := FALSE;
END_VAR

VAR_TEMP
    risingAck : BOOL;
END_VAR

// Detect rising edge of ackBtn
risingAck := ackBtn AND NOT prev_ackBtn;

// Alarm state machine
IF flowLow THEN
    // Condition is active
    IF NOT alarmActive THEN
        // New alarm activation
        alarmActive := TRUE;
        alarmAcked  := FALSE;
    ELSIF risingAck THEN
        // Acknowledge while condition still exists
        alarmAcked := TRUE;
    END_IF;
ELSE
    // Condition has disappeared
    IF alarmActive AND NOT alarmAcked THEN
        // Unacknowledged alarm - enter pending clear state
        alarmAcked := TRUE;
    ELSIF alarmActive AND alarmAcked AND risingAck THEN
        // Acknowledged alarm with condition cleared - clear alarm
        alarmActive := FALSE;
        alarmAcked  := FALSE;
    END_IF;
END_IF;

// High priority alarm: sensor failure (independent of low priority alarm)
highHigh := NOT sensorOK;

// Update state for next cycle
prev_flowLow    := flowLow;
prev_ackBtn     := ackBtn;
prev_alarmAcked := alarmAcked;

END_FUNCTION_BLOCK

(* ---- self-hard-01.candidate_02.st ---- *)
FUNCTION_BLOCK FB
VAR_INPUT
    flowLow   : BOOL;
    ackBtn    : BOOL;
    sensorOK  : BOOL;
END_VAR
VAR_OUTPUT
    alarmActive : BOOL;
    alarmAcked  : BOOL;
    highHigh    : BOOL;
END_VAR
VAR
    prev_flowLow : BOOL := FALSE;
    prev_ackBtn  : BOOL := FALSE;
END_VAR

VAR_TEMP
    risingAck : BOOL;
END_VAR

risingAck := ackBtn AND NOT prev_ackBtn;

IF flowLow THEN
    // Condition is active
    IF NOT alarmActive THEN
        // New alarm activation
        alarmActive := TRUE;
        alarmAcked  := FALSE;
    ELSIF risingAck THEN
        // Rising ack while condition still exists - just mark acknowledged
        alarmAcked := TRUE;
    END_IF;
ELSE
    // Condition has disappeared
    IF prev_flowLow AND alarmAcked THEN
        // Condition just cleared, was already acknowledged - clear immediately
        alarmActive := FALSE;
        alarmAcked  := FALSE;
    ELSIF prev_flowLow AND NOT alarmAcked THEN
        // Condition just cleared, unacknowledged - enter pending clear state
        alarmAcked := TRUE;
    ELSIF risingAck AND alarmAcked THEN
        // Condition still gone from before, pending clear - clear on new ack
        alarmActive := FALSE;
        alarmAcked  := FALSE;
    END_IF;
END_IF;

// High priority alarm: sensor failure (independent)
highHigh := NOT sensorOK;

// Update state for next cycle
prev_flowLow := flowLow;
prev_ackBtn  := ackBtn;

END_FUNCTION_BLOCK

(* ---- self-hard-01.raw_candidate_01.st ---- *)
FUNCTION_BLOCK FB
VAR_INPUT
    flowLow   : BOOL;
    ackBtn    : BOOL;
    sensorOK  : BOOL;
END_VAR
VAR_OUTPUT
    alarmActive : BOOL;
    alarmAcked  : BOOL;
    highHigh    : BOOL;
END_VAR
VAR
    prev_flowLow   : BOOL := FALSE;
    prev_ackBtn    : BOOL := FALSE;
    prev_alarmAcked : BOOL := FALSE;
END_VAR

VAR_TEMP
    risingAck : BOOL;
END_VAR

// Detect rising edge of ackBtn
risingAck := ackBtn AND NOT prev_ackBtn;

// Alarm state machine
IF flowLow THEN
    // Condition is active
    IF NOT alarmActive THEN
        // New alarm activation
        alarmActive := TRUE;
        alarmAcked  := FALSE;
    ELSIF risingAck THEN
        // Acknowledge while condition still exists
        alarmAcked := TRUE;
    END_IF;
ELSE
    // Condition has disappeared
    IF alarmActive AND NOT alarmAcked THEN
        // Unacknowledged alarm - enter pending clear state
        alarmAcked := TRUE;
    ELSIF alarmActive AND alarmAcked AND risingAck THEN
        // Acknowledged alarm with condition cleared - clear alarm
        alarmActive := FALSE;
        alarmAcked  := FALSE;
    END_IF;
END_IF;

// High priority alarm: sensor failure (independent of low priority alarm)
highHigh := NOT sensorOK;

// Update state for next cycle
prev_flowLow    := flowLow;
prev_ackBtn     := ackBtn;
prev_alarmAcked := alarmAcked;

END_FUNCTION_BLOCK
